(* IEC 61131-3 sources: Antarbhukti-LLM/DatasetCreation/SeedSTs/batch1_filtered_BASIC (part 2) *)

(* ---- FT_PROFILE.ST ---- *)
(*@PROPERTIES_EX@
TYPE: POU
LOCALE: 0
IEC_LANGUAGE: ST
PLC_TYPE: independent
PROC_TYPE: independent
GROUP: ENGINEERING.AUTOMATION
*)
(*@KEY@:DESCRIPTION*)
version 1.1	15 sep 2007
programmer 	tobias
tested by	hugo

FT_Profile generates an output signal which is defined by values over a time scale.
the different values are connected by ramps between the individual values.
a rising edge on E starts the output signal generation and E = True can delay time_3 / value_3 as long as it stays true.
an additional multiplier K can be used to multiply the output and an offset O can be added to the output dynamically.
(*@KEY@:END_DESCRIPTION*)
FUNCTION_BLOCK FT_PROFILE

(*Group:Default*)

VAR_INPUT
	K :	REAL := 1.0;
	O :	REAL := 0.0;
	M :	REAL := 1.0;
	E :	BOOL;
	VALUE_0 :	REAL;
	TIME_1 :	TIME;
	VALUE_1 :	REAL;
	TIME_2 :	TIME;
	VALUE_2 :	REAL;
	TIME_3 :	TIME;
	VALUE_3 :	REAL;
	TIME_10 :	TIME;
	VALUE_10 :	REAL;
	TIME_11 :	TIME;
	VALUE_11 :	REAL;
	TIME_12 :	TIME;
	VALUE_12 :	REAL;
	TIME_13 :	TIME;
	VALUE_13 :	REAL;
END_VAR

VAR_OUTPUT
	Y :	REAL;
	RUN :	BOOL;
	ET :	TIME;
END_VAR

VAR
	tx :	TIME;
	edge :	BOOL;
	state :	INT;
	ta :	TIME;
	tb :	TIME;
	t0 :	TIME;
	temp :	REAL;
	va :	REAL;
	vb :	REAL;
	T_PLC_MS :	T_PLC_MS;
END_VAR

(*@KEY@: WORKSHEET
NAME: FT_PROFILE
IEC_LANGUAGE: ST
*)
(* read system time *)
T_PLC_MS();
tx:= UDINT_TO_TIME(T_PLC_MS.T_PLC_MS);

(* determine start condition *)
IF E AND NOT edge THEN
	RUN := TRUE;
	ET := t#0s;
	t0 := tx;
	ta := tx;
	tb := multime(time_1, M);
	va := value_0;
	vb := value_1;
	temp := value_0;
	state := 1;
END_IF;
edge := E;

(* generate startup profile *)
IF run THEN
	CASE state OF
		1:	IF tx - ta >= tb THEN
				ta := ta + tb;
				tb := multime(time_2 - time_1, M);
				va := value_1;
				vb := value_2;
				temp := value_1;
				state := 2;
			ELSE
				temp := ((vb - va) * TIME_TO_REAL(tx - ta) / TIME_TO_REAL(tb) + va);
			END_IF;
		2:	IF tx - ta >= tb THEN
				ta := ta + tb;
				tb := multime(time_3 - time_2, M);
				va := value_2;
				vb := value_3;
				temp := value_2;
				state := 3;
			ELSE
				temp := ((vb - va) * TIME_TO_REAL(tx - ta) / TIME_TO_REAL(tb) + va);
			END_IF;
		3:	IF tx - ta >= tb THEN
				ta := ta + tb;
				tb := multime(time_10 - time_3, M);
				va := value_3;
				vb := value_10;
				temp := value_3;
				state := 4;
			ELSE
				temp := ((vb - va) * TIME_TO_REAL(tx - ta) / TIME_TO_REAL(tb) + va);
			END_IF;
		4 :	IF tx - ta >= tb THEN
				ta := ta + tb;
				tb := multime(time_11 - time_10, M);
				va := value_10;
				vb := value_11;
				temp := value_10;
				IF E THEN state := 5; ELSE state := 6; END_IF;
			ELSE
				temp := ((vb - va) * TIME_TO_REAL(tx - ta) / TIME_TO_REAL(tb) + va);
			END_IF;
		5:	(* extend the signal while E is true *)
			IF E THEN
				ta := tx;
			ELSE
				state := 6;
			END_IF;
		6:	IF tx - ta >= tb THEN
				ta := ta + tb;
				tb := multime(time_12 - time_11, M);
				va := value_11;
				vb := value_12;
				temp := value_11;
				state := 7;
			ELSE
				temp := ((vb - va) * TIME_TO_REAL(tx - ta) / TIME_TO_REAL(tb) + va);
			END_IF;
		7:	IF tx - ta >= tb THEN
				ta := ta + tb;
				tb := multime(time_13 - time_12, M);
				va := value_12;
				vb := value_13;
				temp := value_12;
				state := 8;
			ELSE
				temp := ((vb - va) * TIME_TO_REAL(tx - ta) / TIME_TO_REAL(tb) + va);
			END_IF;
		8:	IF tx - ta >= tb THEN
				temp := value_13;
				run := FALSE;
			ELSE
				temp := ((vb - va) * TIME_TO_REAL(tx - ta) / TIME_TO_REAL(tb) + va);
			END_IF;
	END_CASE;
	Y := temp * K + O;
	ET := tx - t0;
END_IF;

(* revision history
hm	27 feb 2007		rev 1.0
	original version

hm	15. sep2007		rev 1.1
	replaced Time() with T_PLC_MS for compatibility and performance reasons

*)
(*@KEY@: END_WORKSHEET *)
END_FUNCTION_BLOCK

(* ---- FT_PT1.ST ---- *)
(*@PROPERTIES_EX@
TYPE: POU
LOCALE: 0
IEC_LANGUAGE: ST
PLC_TYPE: independent
PROC_TYPE: independent
GROUP: ENGINEERING.CONTROL
*)
(*@KEY@:DESCRIPTION*)
version 1.11	18. jan. 2011
programmer 		hugo
tested by		oscat

FT_PT1 is an low pass filter with a programmable time T and faktor K.

(*@KEY@:END_DESCRIPTION*)
FUNCTION_BLOCK FT_PT1

(*Group:Default*)

VAR_INPUT
	IN :	REAL;
	T :	TIME;
	K :	REAL := 1.0;
END_VAR

VAR_OUTPUT
	OUT :	REAL;
END_VAR

VAR
	last :	UDINT;
	tx :	UDINT;
	init :	BOOL;
	T_PLC_US :	T_PLC_US;
END_VAR

(*@KEY@: WORKSHEET
NAME: FT_PT1
IEC_LANGUAGE: ST
*)
(* read system time *)
T_PLC_US();
tx:= T_PLC_US.T_PLC_US;

(* startup initialisation *)
IF NOT init OR T = t#0s THEN
	init := TRUE;
	out := K * in;
ELSE
	out := out + (in * K - out) * UDINT_TO_REAL(Tx - last) / TIME_TO_REAL(T) * 1.0E-3;
	IF ABS(out) < 1.0E-20 THEN out := 0.0; END_IF;
END_IF;
last := tx;

(*
hm 1.1.2007	rev 1.1
	corrected error while startup value was not correct
	for very small time values real output would run out of range.

hm 3.1.2007	rev 1.2
	corrected an error for falling edge failures.
	added output faktor K.

hm 27. 2. 2007	rev 1.3
	output will be input during init for definitive startup condition.

hm	15.9.2007	rev 1.4
	changed time() to T_PLC_US() for compatibilitxy resons
	increased internal accuracy to Microseconds instead of Milliseconds

hm	23. oct 2007	rev 1.5
	added out := in to the init statements

hm	30. nov 2007	rev 1.6
	changed out to be K * in during initialization

hm	5. jan 2008	rev 1.7
	improved code for better performance

hm	16. mar. 2008	rev 1.8
	added type conversion to avoid warning under codesys 3.0

hm	14. jun. 2008	rev 1.9
	improved code

hm	11. mar. 2009	rev 1.10
	real constants updated to new systax using dot

hm	18. jan. 2011	rev 1.11
	avoid underrun of out
*)
(*@KEY@: END_WORKSHEET *)
END_FUNCTION_BLOCK

(* ---- FT_PT2.ST ---- *)
(*@PROPERTIES_EX@
TYPE: POU
LOCALE: 0
IEC_LANGUAGE: ST
PLC_TYPE: independent
PROC_TYPE: independent
GROUP: ENGINEERING.CONTROL
*)
(*@KEY@:DESCRIPTION*)
version 1.5	11. mar. 2009
programmer 	hugo
tested by	oscat

FT_PT2 is a 2nd grade filter with programmable times T, D and faktor K.
(*@KEY@:END_DESCRIPTION*)
FUNCTION_BLOCK FT_PT2

(*Group:Default*)

VAR_INPUT
	IN :	REAL;
	T :	TIME;
	D :	REAL;
	K :	REAL := 1.0;
END_VAR

VAR_OUTPUT
	OUT :	REAL;
END_VAR

VAR
	init :	BOOL;
	int1 :	INTEGRATE;
	int2 :	INTEGRATE;
	tn :	REAL;
	I1 :	REAL;
	I2 :	REAL;
	tn2 :	REAL;
END_VAR

(*@KEY@: WORKSHEET
NAME: FT_PT2
IEC_LANGUAGE: ST
*)
(* startup initialisation *)
IF NOT init OR T = T#0s THEN
	init := TRUE;
	out := K * in;
	I2 := out;
ELSE
	TN := TIME_TO_REAL(T) / 1000.0;
	tn2 := TN * TN;
	int1(X := in * K / tn2 - I1 * 0.5 * D / TN - I2 / TN2, Y := I1);
	I1 := int1.Y;
	int2(X := I1,Y := I2);
	I2 := int2.Y;
	out := I2;
END_IF;

(* revision history

15.1.2007 hm		rev 1.1
	changed formula to new more acurate formula

hm 15.9.2007		rev 1.2
	deleted unused code for init system time reading tx

hm	30.11.2007	rev 1.3
	changed out to be K * in during initialization
	avoind divide by 0 if tn = 0

hm	3. nov. 2008	rev 1.4
	optimized code and fixed a problem with init

hm	11. mar. 2009	rev 1.5
	real constants updated to new systax using dot

*)
(*@KEY@: END_WORKSHEET *)
END_FUNCTION_BLOCK

(* ---- FT_RMP.ST ---- *)
(*@PROPERTIES_EX@
TYPE: POU
LOCALE: 0
IEC_LANGUAGE: ST
PLC_TYPE: independent
PROC_TYPE: independent
GROUP: MATHEMATICAL.FUNCTIONS
*)
(*@KEY@:DESCRIPTION*)
version 1.4	25 jan 2008
programmer 	oscat
tested BY	oscat

this ramp function follows an input signal with a linear ramp up or down, the up or down speed can be set with KF and KR.
a K factor of 1 means 1 unit per second on the output. K factors can only be positive and not negative.
a busy output signals the ramp is running or busy false means the in value is present on the output.
a rmp input false means the output follows the input dierctly while a rmp = true means the output follows the input with a ramp.
a updn output signal the directon of the ramp (up or down).
(*@KEY@:END_DESCRIPTION*)
FUNCTION_BLOCK FT_RMP

(*Group:Default*)

VAR_INPUT
	RMP :	BOOL := TRUE;
	IN :	REAL;
	KR :	REAL;
	KF :	REAL;
END_VAR

VAR_OUTPUT
	OUT :	REAL;
	BUSY :	BOOL;
	UD :	BOOL;
END_VAR

VAR
	tx :	TIME;
	last :	TIME;
	init :	BOOL;
	T_PLC_MS :	T_PLC_MS;
END_VAR

(*@KEY@: WORKSHEET
NAME: FT_RMP
IEC_LANGUAGE: ST
*)
(* read system time *)
T_PLC_MS();
tx:= UDINT_TO_TIME(T_PLC_MS.T_PLC_MS) - last;

IF NOT init THEN
	init := TRUE;
	last := tx;
	tx := t#0s;
	out := in;
END_IF;
IF NOT rmp THEN
	out := in;
	busy := FALSE;
ELSIF out > in THEN
	(* ramp down *)
	out := out - TIME_TO_REAL(tx) * 0.001 * KF;
	out := MAX(in, out);
ELSIF out < in THEN
	(* ramp up *)
	out := out + TIME_TO_REAL(tx) * 0.001 * KR;
	out := MIN(in, out);
END_IF;

(* set busy and dir flags *)
IF out < in THEN
	busy := TRUE;
	ud := TRUE;
ELSIF out > in THEN
	busy := TRUE;
	ud := FALSE;
ELSE
	busy := FALSE;
END_IF;
last := last + tx;

(* revision history:

hm 8.10.2006			rev 1.1
	added ud output

hm 12. feb 2007		rev 1.2
	added init variable and corrected a possible startup problem

hm	17. sep 2007	rev 1.3
	replaced time() with t_plc_ms() for compatibility reasons

hm	25. jan 2008	rev 1.4
	performance improvements
	allow KR and KF to be 0
*)
(*@KEY@: END_WORKSHEET *)
END_FUNCTION_BLOCK

(* ---- GEN_PULSE.ST ---- *)
(*@PROPERTIES_EX@
TYPE: POU
LOCALE: 0
IEC_LANGUAGE: ST
PLC_TYPE: independent
PROC_TYPE: independent
GROUP: ENGINEERING.SIGNAL_GENERATORS
*)
(*@KEY@:DESCRIPTION*)
version 1.5	8. apr. 2011
programmer 	hugo
tested by	oscat

GEN_PULSE uses the internal sps timer to generate a continuous output waveform with programmable high and low time.
the accuracy of gen_pulse is depending on the system timer.
when time is 0 the high and low times are exactly one cycle.
ENQ = TRUE will start and ENQ = FALSE will stop the generator.
(*@KEY@:END_DESCRIPTION*)
FUNCTION_BLOCK GEN_PULSE

(*Group:Default*)

VAR_INPUT
	ENQ :	BOOL := TRUE;
	PTH :	TIME;
	PTL :	TIME;
END_VAR

VAR_OUTPUT
	Q :	BOOL;
END_VAR

VAR
	T_PLC_MS :	T_PLC_MS;
	tx :	TIME;
	tn :	TIME;
	init :	BOOL;
END_VAR

(*@KEY@: WORKSHEET
NAME: GEN_PULSE
IEC_LANGUAGE: ST
*)
IF enq THEN
	T_PLC_MS();	(* read system timer *)
	tx:= UDINT_TO_TIME(T_PLC_MS.T_PLC_MS);
	IF NOT init THEN init := TRUE; tn := tx; END_IF;
	IF tx - tn >= SEL(Q, PTL, PTH) THEN
		tn := tn + SEL(Q, PTL, PTH);
		Q := NOT Q;
	END_IF;
ELSE
	Q := FALSE;
	init := FALSE;
END_IF;

(* revision history
hm	29. jun. 2008	rev 1.0
	original version

hm	23. nov. 2008	rev 1.1
	set default for enq to be true

hm	18. jul. 2009	rev 1.2
	improved performance

hm	13. nov. 2009	rev 1.3
	corrected error

hm	16. feb. 2011	rev 1.4
	corrected an error when timer overflows

hm	8. apr. 2011	rev 1.5
	ptl and pth was exchanged
*)
(*@KEY@: END_WORKSHEET *)
END_FUNCTION_BLOCK

(* ---- GEN_RMP.ST ---- *)
(*@PROPERTIES_EX@
TYPE: POU
LOCALE: 0
IEC_LANGUAGE: ST
PLC_TYPE: independent
PROC_TYPE: independent
GROUP: ENGINEERING.SIGNAL_GENERATORS
*)
(*@KEY@:DESCRIPTION*)
version 1.4	10. mar. 2009
programmer 	oscat
tested BY	oscat

this signal generator generates a ramp wave output. The ramp wave signal is defined by period time (PT),
amplitude (AM), offset (OS) and a specific delay for the output signal (DL).
The Output waveform will have its minimum peak at OS and its maximum peak at AM + OS.
The delay input can delay a signal up to PT, this can be useful to synchronize different generators
and generate interleaving signals.
in addition to the analog output Out there is a second boolean output Q with is true for one cycle when the ramp starts.

(*@KEY@:END_DESCRIPTION*)
FUNCTION_BLOCK GEN_RMP

(*Group:Default*)

VAR_INPUT
	PT :	TIME := T#1s;
	AM :	REAL := REAL#1.0;
	OS :	REAL;
	DL :	REAL;
END_VAR

VAR_OUTPUT
	Q :	BOOL;
	OUT :	REAL;
END_VAR

VAR
	tx :	TIME;
	last :	TIME;
	init :	BOOL;
	temp :	REAL;
	ltemp :	REAL;
	T_PLC_MS :	T_PLC_MS;
END_VAR

(*@KEY@: WORKSHEET
NAME: GEN_RMP
IEC_LANGUAGE: ST
*)
(* read system time and prepare input data *)
T_PLC_MS();
tx:= UDINT_TO_TIME(T_PLC_MS.T_PLC_MS) - last;
DL := modR(dl,1.0);
IF dl < 0.0 THEN dl := 1.0 - dl; END_IF;

(* init section *)
IF NOT init THEN
	init := TRUE;
	last := tx;
	tx := t#0s;
END_IF;

(* add last if one cycle is finished *)
IF tx >= pt THEN
	last := last + pt;
	tx := tx - pt;
END_IF;

(* generate sine wave *)
ltemp := temp;
IF pt > t#0s THEN temp := fract(TIME_TO_REAL(tx + multime(pt, dl)) / TIME_TO_REAL(pt)); END_IF;
out := am * temp + os;

(* boolean output Q *)
Q := temp < ltemp;

(* revision history
hm	3. mar 2007		rev 1.0
	original version

hm	17 sep 2007		rev 1.1
	replaced time() with t_plc_ms for compatibilitx reasons

hm	27. nov 2007	rev 1.2
	avoid divide by 0 when pt = 0

ks	26. oct. 2008	rev 1.3
	code optimization

hm	10. mar. 2009	rev 1.4
	changed real constants to use dot syntax
*)
(*@KEY@: END_WORKSHEET *)
END_FUNCTION_BLOCK

(* ---- GEN_SQ.ST ---- *)
(*@PROPERTIES_EX@
TYPE: POU
LOCALE: 0
IEC_LANGUAGE: ST
PLC_TYPE: independent
PROC_TYPE: independent
GROUP: LOGIC.GENERATORS
*)
(*@KEY@:DESCRIPTION*)
version 1.3	16. feb. 2011
programmer 	    hugo
tested by		tobias

gen_sq generates square wave signal with programmable period time.

(*@KEY@:END_DESCRIPTION*)
FUNCTION_BLOCK GEN_SQ

(*Group:Default*)

VAR_INPUT
	PT :	TIME;
END_VAR

VAR_OUTPUT
	Q :	BOOL;
END_VAR

VAR
	init :	BOOL;
	tn :	TIME;
	tx :	TIME;
	T_PLC_MS :	T_PLC_MS;
END_VAR

(*@KEY@: WORKSHEET
NAME: GEN_SQ
IEC_LANGUAGE: ST
*)
(* read system time *)
T_PLC_MS();
tx := UDINT_TO_TIME(T_PLC_MS.T_PLC_MS);

IF NOT init THEN
	init := TRUE;
	tn := tx;
	Q := TRUE;
ELSIF tx - tn >= DWORD_TO_TIME(SHR(TIME_TO_DWORD(PT),1)) THEN
	Q := NOT Q;
	tn := tn + DWORD_TO_TIME(SHR(TIME_TO_DWORD(pt),1));
END_IF;

(* revision history
hm	4. aug 2006	rev 1.0
	original version

hm	17. sep 2007	rev 1.1
	replaced time() with T_PLC_MS() for compatibility reasons

hm	18. jul. 2009	rev 1.2
	improved accuracy

hm	16. feb 2011	rev 1.3
	corrected an error with timer overflow
*)

(*@KEY@: END_WORKSHEET *)
END_FUNCTION_BLOCK

(* ---- HYST.ST ---- *)
(*@PROPERTIES_EX@
TYPE: POU
LOCALE: 0
IEC_LANGUAGE: ST
PLC_TYPE: independent
PROC_TYPE: independent
GROUP: ENGINEERING.CONTROL
*)
(*@KEY@:DESCRIPTION*)
version 1.0	2. jun. 2008
programmer 	hugo
tested BY	tobias

This Hystereses function has two modes:
1. if on > off then Q will be switched high when in > on and switched low when in < off.
2. if on < off then Q will be switched high when in < on and switched low when in > off.
the output win will be high when in is between low and high.
(*@KEY@:END_DESCRIPTION*)
FUNCTION_BLOCK HYST

(*Group:Default*)

VAR_INPUT
	IN :	REAL;
	ON :	REAL;
	OFF :	REAL;
END_VAR

VAR_OUTPUT
	Q :	BOOL;
	WIN :	BOOL;
END_VAR

(*@KEY@: WORKSHEET
NAME: HYST
IEC_LANGUAGE: ST
*)
IF ON >= OFF THEN
	IF IN < OFF THEN
		Q := FALSE;
		WIN := FALSE;
	ELSIF  IN > ON THEN
		Q := TRUE;
		WIN := FALSE;
	ELSE
		WIN := TRUE;
	END_IF;
ELSE
	IF IN > OFF THEN
		Q := FALSE;
		WIN := FALSE;
	ELSIF  IN < ON THEN
		Q := TRUE;
		WIN := FALSE;
	ELSE
		WIN := TRUE;
	END_IF;
END_IF;

(* revision history
hm		2.  jun 2008	rev 1.0
	original version

*)
(*@KEY@: END_WORKSHEET *)
END_FUNCTION_BLOCK

(* ---- HYST_1.ST ---- *)
(*@PROPERTIES_EX@
TYPE: POU
LOCALE: 0
IEC_LANGUAGE: ST
PLC_TYPE: independent
PROC_TYPE: independent
GROUP: ENGINEERING.CONTROL
*)
(*@KEY@:DESCRIPTION*)
version 1.1	2. jun. 2008
programmer 	hugo
tested BY	tobias

this hysteresis function switches the output high if the input signal reaches obove high and will switch to low when the input falls back below low value.
a separate output mid is set if the input stays between low and high value.
(*@KEY@:END_DESCRIPTION*)
FUNCTION_BLOCK HYST_1

(*Group:Default*)

VAR_INPUT
	IN :	REAL;
	HIGH :	REAL;
	LOW :	REAL;
END_VAR

VAR_OUTPUT
	Q :	BOOL;
	WIN :	BOOL;
END_VAR

(*@KEY@: WORKSHEET
NAME: HYST_1
IEC_LANGUAGE: ST
*)
IF in < low THEN
	Q := FALSE;
	win := FALSE;
ELSIF in > high THEN
	Q := TRUE;
	win := FALSE;
ELSE
	win := TRUE;
END_IF;

(* code used for rev 1.0
IF Q THEN
	IF in < low THEN q := FALSE; END_IF;
ELSE
	IF in > high THEN q := TRUE; END_IF;
END_IF;
win := in > low AND in < high;
*)
(*@KEY@: END_WORKSHEET *)
END_FUNCTION_BLOCK

(* ---- HYST_2.ST ---- *)
(*@PROPERTIES_EX@
TYPE: POU
LOCALE: 0
IEC_LANGUAGE: ST
PLC_TYPE: independent
PROC_TYPE: independent
GROUP: ENGINEERING.CONTROL
*)
(*@KEY@:DESCRIPTION*)
version 1.2	2. jun. 2008
programmer 	oscat
tested BY	tobias

this hysteresis function switches the output high if the input signal reaches obove val + hys/2 and will switch to low when the input falls back below val - hys/2 value.
a separate output mid is set if the input stays between low and high value.
(*@KEY@:END_DESCRIPTION*)
FUNCTION_BLOCK HYST_2

(*Group:Default*)

VAR_INPUT
	IN :	REAL;
	VAL :	REAL;
	HYS :	REAL;
END_VAR

VAR_OUTPUT
	Q :	BOOL;
	WIN :	BOOL;
END_VAR

VAR
	tmp :	REAL;
END_VAR

(*@KEY@: WORKSHEET
NAME: HYST_2
IEC_LANGUAGE: ST
*)
tmp := val - hys * 0.5;
IF in < tmp THEN
	Q := FALSE;
	win := FALSE;
ELSIF in > tmp + hys THEN
	Q := TRUE;
	win := FALSE;
ELSE
	win := TRUE;
END_IF;

(* code used for 1.2 and before
X := hys * 0.5;
IF Q THEN
	IF in < val - x THEN q := FALSE; END_IF;
ELSE
	IF in > val + x THEN q := TRUE; END_IF;
END_IF;
win := in > val - x AND in < val + x;
*)

(* revision history
hm		4. aug 2006	rev 1.0
	original version

hm		5. jan 2008	rev 1.1
	improved code for better performance

hm		2. jun. 2008	rev 1.2
	improved performance
*)
(*@KEY@: END_WORKSHEET *)
END_FUNCTION_BLOCK

(* ---- HYST_3.ST ---- *)
(*@PROPERTIES_EX@
TYPE: POU
LOCALE: 0
IEC_LANGUAGE: ST
PLC_TYPE: independent
PROC_TYPE: independent
GROUP: ENGINEERING.CONTROL
*)
(*@KEY@:DESCRIPTION*)
version 1.2	5 jan 2008
programmer 	oscat
tested BY	tobias

this is a double hysteresis function. Out1 follows a hysteresis function defined by val1and hyst, while out 2 follows val2 and hyst.
if the input signal is between the two hysteresis switches (val1 and val2) then non of the outputs is active.
(*@KEY@:END_DESCRIPTION*)
FUNCTION_BLOCK HYST_3

(*Group:Default*)

VAR_INPUT
	IN :	REAL;
	HYST :	REAL;
	VAL1 :	REAL;
	VAL2 :	REAL;
END_VAR

VAR_OUTPUT
	Q1 :	BOOL;
	Q2 :	BOOL;
END_VAR

VAR
	X :	REAL;
END_VAR

(*@KEY@: WORKSHEET
NAME: HYST_3
IEC_LANGUAGE: ST
*)
X := hyst * 0.5;
IF in < val1 - X THEN
	q1 := TRUE;
ELSIF in > val1 + X THEN
	q1 := FALSE;
END_IF;
IF in < val2 - X THEN
	q2 := FALSE;
ELSIF in > val2 + X THEN
	q2 := TRUE;
END_IF;

(* revision history
hm	22. jan 2007	rev 1.0
	original version

hm	27. dec 2007	rev 1.1
	changed code for better performance

hm	5. jan 2008		rev 1.2
	further performance iprovements

*)
(*@KEY@: END_WORKSHEET *)
END_FUNCTION_BLOCK

(* ---- INC_DEC.ST ---- *)
(*@PROPERTIES_EX@
TYPE: POU
LOCALE: 0
IEC_LANGUAGE: ST
PLC_TYPE: independent
PROC_TYPE: independent
GROUP: ENGINEERING.AUTOMATION
*)
(*@KEY@:DESCRIPTION*)
version 1.0	4 aug 2006
programmer 	oscat
tested BY	oscat

incremental decoder with quadruple accuracy.
2 pulses for each channel are created for each directional pulse.
(*@KEY@:END_DESCRIPTION*)
FUNCTION_BLOCK INC_DEC

(*Group:Default*)

VAR_INPUT
	CHA :	BOOL;
	CHB :	BOOL;
	RST :	BOOL := 0;
END_VAR

VAR_OUTPUT
	DIR :	BOOL;
	CNT :	INT;
END_VAR

VAR
	edgea :	BOOL := 0;
	clk :	BOOL;
	clka :	BOOL;
	clkb :	BOOL;
	edgeb :	BOOL;
	axb :	BOOL;
END_VAR

(*@KEY@: WORKSHEET
NAME: INC_DEC
IEC_LANGUAGE: ST
*)
axb := cha XOR chb;

(* create pulses for channel a *)
clka := cha XOR edgea;
edgea := cha;

clkb := chb XOR edgeb;
edgeb := chb;

(* create pulses for both channels *)
clk := clka OR clkb;

(* set the direction output *)
IF axb AND clka THEN dir := TRUE; END_IF;
IF axb AND clkb THEN dir := FALSE; END_IF;

(* increment or decrement the counter *)
IF clk AND dir THEN cnt := cnt + 1; END_IF;
IF clk AND NOT dir THEN cnt := cnt -1; END_IF;

(* reset the counter if rst active *)
IF rst THEN cnt := 0; END_IF;
(*@KEY@: END_WORKSHEET *)
END_FUNCTION_BLOCK

(* ---- INTERLOCK.ST ---- *)
(*@PROPERTIES_EX@
TYPE: POU
LOCALE: 0
IEC_LANGUAGE: ST
PLC_TYPE: independent
PROC_TYPE: independent
GROUP: ENGINEERING.AUTOMATION
*)
(*@KEY@:DESCRIPTION*)
version 1.0	28 sep 2007
programmer 	hugo
tested by	tobias

INTERLOCK has two inputs I1 and I2 which drive the corresponding outputs Q1 and Q2.
the inputs signals lock each other out and therfore I1 can only drive Q1 when I2 is Low and vice versa.
The input TL specifies a dead time between two outputs can become active.
an output can only become active when the other output was not active for the time TL.
(*@KEY@:END_DESCRIPTION*)
FUNCTION_BLOCK INTERLOCK

(*Group:Default*)

VAR_INPUT
	I1 :	BOOL;
	I2 :	BOOL;
	TL :	TIME;
END_VAR

VAR_OUTPUT
	Q1 :	BOOL;
	Q2 :	BOOL;
END_VAR

VAR
	T1 :	TOF;
	T2 :	TOF;
END_VAR

(*@KEY@: WORKSHEET
NAME: INTERLOCK
IEC_LANGUAGE: ST
*)
(* the input signal have a run delay to lockout the other input *)
T1(IN := I1, PT := TL);
T2(IN := I2, PT := TL);

Q1 := I1 AND NOT t2.Q;
Q2 := I2 AND NOT t1.Q;

(* revision history

hm	28 sep 2007		rev 1.0
	original version

*)
(*@KEY@: END_WORKSHEET *)
END_FUNCTION_BLOCK

(* ---- INTERLOCK_4.ST ---- *)
(*@PROPERTIES_EX@
TYPE: POU
LOCALE: 0
IEC_LANGUAGE: ST
PLC_TYPE: independent
PROC_TYPE: independent
GROUP: ENGINEERING.AUTOMATION
*)
(*@KEY@:DESCRIPTION*)
version 1.1	14. mar. 2009
programmer 	hugo
tested by	oscat

INTERLOCK_4 detects one of 4 switches and delivers the number of the switch pressed on the output out
a output tp is true for one cycle if the output has changed.
a setup variable MODE selects between 3 different modes:
MODE = 0, any input active will disable all other inputs
MODE = 1, the input with the highest number will be acepted
mode = 2, the input last pressed will disable all others

(*@KEY@:END_DESCRIPTION*)
FUNCTION_BLOCK INTERLOCK_4

(*Group:Default*)

VAR_INPUT
	I0 :	BOOL;
	I1 :	BOOL;
	I2 :	BOOL;
	I3 :	BOOL;
	E :	BOOL;
	MODE :	INT;
END_VAR

VAR_OUTPUT
	OUT :	BYTE;
	TP :	BOOL;
END_VAR

VAR
	in :	BYTE;
	last :	BYTE;
	old :	BYTE;
	lmode :	INT;
END_VAR

(*@KEY@: WORKSHEET
NAME: INTERLOCK_4
IEC_LANGUAGE: ST
*)
(* check if enable is active *)
IF E THEN
(* reset all vars when there is a mode change on thy fly *)
	IF mode <> lmode THEN
		out := BYTE#0;
		last := BYTE#0;
		old := BYTE#0;
		lmode := mode;
	END_IF;
	(* load inputs into in *)
	in:=BIT_LOAD_B(in,I0,0); (* in.0 *)
	in:=BIT_LOAD_B(in,I1,1); (* in.1 *)
	in:=BIT_LOAD_B(in,I2,2); (* in.2 *)
	in:=BIT_LOAD_B(in,I3,3); (* in.3 *)
	(* only execute when there is any change *)
	IF in <> last THEN
		(* only execute when inputs have chages state *)
		CASE mode OF
			0:	(* output directly display inputs as bits in byte out *)
				out := in;

			1:	(* the input with the highest number will be acepted *)
				IF    (in AND BYTE#2#00001000) > BYTE#0 (* in.3 *) THEN out := BYTE#8;
				ELSIF (in AND BYTE#2#00000100) > BYTE#0 (* in.2 *) THEN out := BYTE#4;
				ELSIF (in AND BYTE#2#00000010) > BYTE#0 (* in.1 *) THEN out := BYTE#2;
				ELSE out := in;
				END_IF;

			2:	(* input last pressed will be displayed only *)
				last := ((in XOR last) AND in);
				IF    (last AND BYTE#2#00001000) > BYTE#0 (* last.3 *) THEN out := BYTE#8;
				ELSIF (last AND BYTE#2#00000100) > BYTE#0 (* last.2 *) THEN out := BYTE#4;
				ELSIF (last AND BYTE#2#00000010) > BYTE#0 (* last.1 *) THEN out := BYTE#2;
				ELSE out := last;
				END_IF;

			3:	(* any input active will disable all other inputs *)
				IF (out AND in) = BYTE#0 THEN
					IF    (in AND BYTE#2#00001000) > BYTE#0 (* in.3 *) THEN out := BYTE#8;
					ELSIF (in AND BYTE#2#00000100) > BYTE#0 (* in.2 *) THEN out := BYTE#4;
					ELSIF (in AND BYTE#2#00000010) > BYTE#0 (* in.1 *) THEN out := BYTE#2;
					ELSE out := in;
					END_IF;
				END_IF;

		END_CASE;
		last := in;
	END_IF;
	tp := out <> old;
	old := out;
ELSE
	out := BYTE#0;
	last := BYTE#0;
	old := BYTE#0;
	lmode := 0;
	tp := FALSE;
END_IF;

(* revision history
hm	24. oct 2008	rev 1.0
	original version

hm	14. mar. 2009	rev 1.1
	replaced double assignments

*)
(*@KEY@: END_WORKSHEET *)
END_FUNCTION_BLOCK

(* ---- LTCH.ST ---- *)
(*@PROPERTIES_EX@
TYPE: POU
LOCALE: 0
IEC_LANGUAGE: ST
PLC_TYPE: independent
PROC_TYPE: independent
GROUP: LOGIC.FF_PULSE_TRIGGERED
*)
(*@KEY@:DESCRIPTION*)
version 1.2	30. oct. 2008
programmer 	hugo
tested by	oscat

Transparent Latch with asynchronous reset
(*@KEY@:END_DESCRIPTION*)
FUNCTION_BLOCK LTCH

(*Group:Default*)

VAR_INPUT
	D :	BOOL;
	L :	BOOL;
	RST :	BOOL;
END_VAR

VAR_OUTPUT
	Q :	BOOL;
END_VAR

(*@KEY@: WORKSHEET
NAME: LTCH
IEC_LANGUAGE: ST
*)
(* as long as L is true, the latch is transparent and and change of D is transferred to Q *)
(* of course only when there is no asynchronous reset *)
IF rst THEN				(* if asynchronous reset then Q=0 *)
	Q := FALSE;
ELSIF L THEN			(* latch is transparent *)
	Q := D;
END_IF;

(* revision history
hm	4. aug 2006		rev 1.0
	original version

hm	27. dec 2007	rev 1.1
	changed code for better performance

hm	30. oct. 2008	rev 1.2
	deleted unnecessary init with 0

*)
(*@KEY@: END_WORKSHEET *)
END_FUNCTION_BLOCK

(* ---- LTCH_4.ST ---- *)
(*@PROPERTIES_EX@
TYPE: POU
LOCALE: 0
IEC_LANGUAGE: ST
PLC_TYPE: independent
PROC_TYPE: independent
GROUP: LOGIC.FF_PULSE_TRIGGERED
*)
(*@KEY@:DESCRIPTION*)
version 1.3	14. mar. 2009
programmer 	hugo
tested by	oscat

Quad Transparent Latch with asynchronous reset
(*@KEY@:END_DESCRIPTION*)
FUNCTION_BLOCK LTCH_4

(*Group:Default*)

VAR_INPUT
	D0 :	BOOL;
	D1 :	BOOL;
	D2 :	BOOL;
	D3 :	BOOL;
	L :	BOOL;
	RST :	BOOL;
END_VAR

VAR_OUTPUT
	Q0 :	BOOL;
	Q1 :	BOOL;
	Q2 :	BOOL;
	Q3 :	BOOL;
END_VAR

(*@KEY@: WORKSHEET
NAME: LTCH_4
IEC_LANGUAGE: ST
*)
(* as long as L is true, the latch is transparent and and change of D is transferred to Q *)
(* of course only when there is no asynchronous reset *)
IF rst THEN			(* if asynchronous reset then Q=0 *)
	Q0 := FALSE;
	Q1 := FALSE;
	Q2 := FALSE;
	Q3 := FALSE;
ELSIF L THEN			(* latch is transparent *)
	Q0 := D0;
	Q1 := D1;
	Q2 := D2;
	Q3 := D3;
END_IF;

(* revision history
hm	4. aug 2006	rev 1.0
	original version

hm	27. dec 2007	rev 1.1
	changed code for better performance

hm	30. oct. 2008	rev 1.2
	deleted unnecessary init with 0

hm	14. mar. 2009	rev 1.3
	removed double assignments

*)
(*@KEY@: END_WORKSHEET *)
END_FUNCTION_BLOCK

(* ---- MANUAL_1.ST ---- *)
(*@PROPERTIES_EX@
TYPE: POU
LOCALE: 0
IEC_LANGUAGE: ST
PLC_TYPE: independent
PROC_TYPE: independent
GROUP: ENGINEERING.AUTOMATION
*)
(*@KEY@:DESCRIPTION*)
version 1.2	14. mar. 2009
programmer 	hugo
tested by	oscat

MANUAL_1 is a manual override for digital signals.
When MAN = FALSE, the output follows IN and when MAN = TRUE the Output follows M_I.

(*@KEY@:END_DESCRIPTION*)
FUNCTION_BLOCK MANUAL_1

(*Group:Default*)

VAR_INPUT
	IN :	BOOL;
	MAN :	BOOL;
	M_I :	BOOL;
	SET :	BOOL;
	RST :	BOOL;
END_VAR

VAR_OUTPUT
	Q :	BOOL;
	STATUS :	BYTE;
END_VAR

VAR
	S_edge :	BOOL;
	r_edge :	BOOL;
	edge :	BOOL;
END_VAR

(*@KEY@: WORKSHEET
NAME: MANUAL_1
IEC_LANGUAGE: ST
*)
IF NOT man THEN
	Q := IN;
	STATUS := BYTE#100;
	edge := FALSE;
ELSIF NOT s_edge AND set THEN
	Q := TRUE;
	edge := TRUE;
	status := BYTE#101;
ELSIF NOT r_edge AND rst THEN
	Q := FALSE;
	edge := TRUE;
	status := BYTE#102;
ELSIF NOT edge THEN
	Q := M_I;
	status := BYTE#103;
END_IF;

(* remember levels of manual signals *)
s_edge := SET;
r_edge := RST;

(* revision history
hm	17. jun 2008	rev 1.0
	original version

hm	17. oct 2008	rev 1.1
	deleted unnecessary variable m_edge

hm	14. mar. 2009	rev 1.2
	replaced double assignments

*)
(*@KEY@: END_WORKSHEET *)
END_FUNCTION_BLOCK

(* ---- MANUAL_2.ST ---- *)
(*@PROPERTIES_EX@
TYPE: POU
LOCALE: 0
IEC_LANGUAGE: ST
PLC_TYPE: independent
PROC_TYPE: independent
GROUP: ENGINEERING.AUTOMATION
*)
(*@KEY@:DESCRIPTION*)
version 1.0	22. sep. 2008
programmer 	hugo
tested by	oscat

MANUAL_2 is a manual override for boolean signals.
it has static force high and low as well as a manual input.
(*@KEY@:END_DESCRIPTION*)
FUNCTION_BLOCK MANUAL_2

(*Group:Default*)

VAR_INPUT
	IN :	BOOL;
	ENA :	BOOL;
	ON :	BOOL;
	OFF :	BOOL;
	MAN :	BOOL;
END_VAR

VAR_OUTPUT
	Q :	BOOL;
	STATUS :	BYTE;
END_VAR

(*@KEY@: WORKSHEET
NAME: MANUAL_2
IEC_LANGUAGE: ST
*)
IF ena THEN
	IF NOT ON AND NOT OFF THEN
		Q := IN;
		STATUS := BYTE#100;
	ELSIF on AND NOT off THEN
		Q := TRUE;
		STATUS := BYTE#101;
	ELSIF NOT on AND off THEN
		q := FALSE;
		STATUS := BYTE#102;
	ELSE
		Q := MAN;
		STATUS := BYTE#103;
	END_IF;
ELSE
	Q := FALSE;
	STATUS := BYTE#104;
END_IF;

(* revision history
hm	22. sep. 2008		rev 1.0
	original version

*)
(*@KEY@: END_WORKSHEET *)
END_FUNCTION_BLOCK

(* ---- MANUAL_4.ST ---- *)
(*@PROPERTIES_EX@
TYPE: POU
LOCALE: 0
IEC_LANGUAGE: ST
PLC_TYPE: independent
PROC_TYPE: independent
GROUP: ENGINEERING.AUTOMATION
*)
(*@KEY@:DESCRIPTION*)
version 1.0	17. jun 2008
programmer 	hugo
tested by	oscat

MANUAL_4 is a manual override for digital signals.
When MAN = FALSE, the output follows IN and when MAN = TRUE the Output follows M_I.
(*@KEY@:END_DESCRIPTION*)
FUNCTION_BLOCK MANUAL_4

(*Group:Default*)

VAR_INPUT
	I0 :	BOOL;
	I1 :	BOOL;
	I2 :	BOOL;
	I3 :	BOOL;
	MAN :	BOOL;
	STP :	BOOL;
	M0 :	BOOL;
	M1 :	BOOL;
	M2 :	BOOL;
	M3 :	BOOL;
END_VAR

VAR_OUTPUT
	Q0 :	BOOL;
	Q1 :	BOOL;
	Q2 :	BOOL;
	Q3 :	BOOL;
	STATUS :	BYTE;
END_VAR

VAR
	edge :	BOOL;
	pos :	INT;
	tog :	BOOL;
END_VAR

(*@KEY@: WORKSHEET
NAME: MANUAL_4
IEC_LANGUAGE: ST
*)
IF man THEN
	IF NOT TOG THEN
		Q0 := M0;
		Q1 := M1;
		Q2 := M2;
		Q3 := M3;
		STATUS := BYTE#101;
	END_IF;
	IF STP AND NOT edge THEN
		tog := TRUE;
		CASE pos OF
			0:	Q0 := TRUE;
				Q1 := FALSE;
				Q2 := FALSE;
				Q3 := FALSE;
				STATUS := BYTE#110;
			1:	Q0 := FALSE;
				Q1 := TRUE;
				Q2 := FALSE;
				Q3 := FALSE;
				STATUS := BYTE#111;
			2:	Q0 := FALSE;
				Q1 := FALSE;
				Q2 := TRUE;
				Q3 := FALSE;
				STATUS := BYTE#112;
			3:	Q0 := FALSE;
				Q1 := FALSE;
				Q2 := FALSE;
				Q3 := TRUE;
				STATUS := BYTE#113;
		END_CASE;
		pos := INC(pos,1,3);
	END_IF;
ELSE
	Q0 := I0;
	Q1 := I1;
	Q2 := I2;
	Q3 := I3;
	STATUS := BYTE#100;
	tog := FALSE;
	pos := 0;
END_IF;

(* remember status of stp *)
edge := STP;

(* revision history
hm	17. jun 2008		rev 1.0
	original version

*)
(*@KEY@: END_WORKSHEET *)
END_FUNCTION_BLOCK

(* ---- MESSAGE_4R.ST ---- *)
(*@PROPERTIES_EX@
TYPE: POU
LOCALE: 0
IEC_LANGUAGE: ST
PLC_TYPE: independent
PROC_TYPE: independent
GROUP: STRINGS
*)
(*@KEY@:DESCRIPTION*)
version 1.1	27. oct. 2008
programmer 	hugo
tested by	tobias

this function generates a rotation meassage with up to 4 strings.
on each rising edge of EN the next message in line will be displayed.
when EN stays high longer then one cycle, the next message will be displayed automatically after the time T1 is elapsed.
the output MX is the generated message and CX is a counter 0..3 signaling the current message displayed.
the displayed messages are 0 .. MM.
(*@KEY@:END_DESCRIPTION*)
FUNCTION_BLOCK MESSAGE_4R

(*Group:Default*)

VAR_INPUT
	M0 :	STRING;
	M1 :	STRING;
	M2 :	STRING;
	M3 :	STRING;
	MM :	INT := 3;
	ENQ :	BOOL := TRUE;
	CLK :	BOOL := TRUE;
	T1 :	TIME := T#3s;
END_VAR

VAR_OUTPUT
	MX :	STRING;
	MN :	INT;
	TR :	BOOL;
END_VAR

VAR
	timer :	TON;
	edge :	BOOL;
END_VAR

(*@KEY@: WORKSHEET
NAME: MESSAGE_4R
IEC_LANGUAGE: ST
*)
(* check for rising edge on EN *)
TR := FALSE;
IF ENQ THEN
	IF (NOT edge AND clk) OR timer.q THEN
			MN := INC1(MN, MM);
			TR := TRUE;
			timer(in := FALSE);
			CASE MN OF
				0 : MX := M0;
				1 : MX := M1;
				2 : MX := M2;
				3 : MX := M3;
			END_CASE;
	END_IF;
	edge := clk;
	timer( in := CLK, pt := T1);
ELSE
	MX := '';
	MN := 0;
END_IF;

(* revision history
hm	8. oct. 2008	rev 1.0
	original version

hm	27. oct. 2008	rev 1.1
	changed _INC to INC1

*)
(*@KEY@: END_WORKSHEET *)
END_FUNCTION_BLOCK

(* ---- MESSAGE_8.ST ---- *)
(*@PROPERTIES_EX@
TYPE: POU
LOCALE: 0
IEC_LANGUAGE: ST
PLC_TYPE: independent
PROC_TYPE: independent
GROUP: STRINGS
*)
(*@KEY@:DESCRIPTION*)
version 1.1	29. mar. 2008
programmer 	hugo
tested by	tobias

this function generates one out of 4 messages specified by S1 .. S8.
the selected message will be presented at the output M.
In1 has higher priority then In2 which has higher priority then IN3 and in8 has the lowest priority.
(*@KEY@:END_DESCRIPTION*)
FUNCTION_BLOCK MESSAGE_8

(*Group:Default*)

VAR_INPUT
	IN1 :	BOOL;
	IN2 :	BOOL;
	IN3 :	BOOL;
	IN4 :	BOOL;
	IN5 :	BOOL;
	IN6 :	BOOL;
	IN7 :	BOOL;
	IN8 :	BOOL;
	S1 :	STRING;
	S2 :	STRING;
	S3 :	STRING;
	S4 :	STRING;
	S5 :	STRING;
	S6 :	STRING;
	S7 :	STRING;
	S8 :	STRING;
END_VAR

VAR_OUTPUT
	M :	STRING;
END_VAR

(*@KEY@: WORKSHEET
NAME: MESSAGE_8
IEC_LANGUAGE: ST
*)
(* check if an alarm is present if yes set the output M otherwise clear M *)
IF in1 THEN
	M := S1;
ELSIF in2 THEN
	M := S2;
ELSIF in3 THEN
	M := S3;
ELSIF in4 THEN
	M := S4;
ELSIF in5 THEN
	M := S5;
ELSIF in6 THEN
	M := S6;
ELSIF in7 THEN
	M := S7;
ELSIF in8 THEN
	M := S8;
ELSE
	M := '';
END_IF;

(* revision history
hm	26.12.2007		rev 1.0
	original version

hm	29. mar. 2008	rev 1.1
	changed STRING to STRING(STRING_LENGTH)
*)
(*@KEY@: END_WORKSHEET *)
END_FUNCTION_BLOCK

(* ---- METER.ST ---- *)
(*@PROPERTIES_EX@
TYPE: POU
LOCALE: 0
IEC_LANGUAGE: ST
PLC_TYPE: independent
PROC_TYPE: independent
GROUP: ENGINEERING.MEASUREMENTS
*)
(*@KEY@:DESCRIPTION*)
version 1.4	8. mar. 2009
programmer 	oscat
tested BY	oscat

METER measures usage of power or similar values the output MX is the sum of the inputs over time.
MX := sum over time of (I1 * P1 + I2 * P2)/D.
a simple example is the consumption counter for a 2 stage oil burner where stage 1 is 10KW and stage 2 is 20KW.
I1 and I2 decide which value is accounted for, I1 = True only counts P1, I2 is True counts P2
and I1 and I2 is true counts P1 and P2.
the meter can be used for all kind of consumption meters. P1 and P2 can change on the fly.

(*@KEY@:END_DESCRIPTION*)
FUNCTION_BLOCK METER

(*Group:Default*)

VAR_INPUT
	M1 :	REAL;
	M2 :	REAL;
	I1 :	BOOL;
	I2 :	BOOL;
	D :	REAL := 1.0;
	RST :	BOOL;
END_VAR

VAR_IN_OUT
	MX :	REAL;
END_VAR

VAR RETAIN
	MR :	REAL2;
END_VAR

VAR
	MX1 :	REAL;(*current consumption value on M1 and M2*)
	MX2 :	REAL;(*current consumption value on M1 and M2*)
	tx :	UDINT;
	last :	UDINT;
	tc :	REAL;
	init :	BOOL;
	T_PLC_MS :	T_PLC_MS;
	R2_ADD :	R2_ADD;
END_VAR

(*@KEY@: WORKSHEET
NAME: METER
IEC_LANGUAGE: ST
*)
(* measure the last cycle time and make sure we onle execute once every millisecond *)
T_PLC_MS();
tx:= T_PLC_MS.T_PLC_MS;
IF NOT init THEN
	init := TRUE;
	last := tx;
	mr.RX := mx;
	mr.R1 := 0.0;
ELSIF tx = last THEN
	RETURN;
ELSE
	tc := UDINT_TO_REAL(tx - last) * 0.001;
END_IF;
last := tx;

(* reset *)
IF rst THEN
	mr.R1 := 0.0;
	mr.RX := 0.0;
ELSE
	(* current consumption measurement *)
	MX1 := SEL(I1,0.0,M1);
	MX2 := SEL(I2,0.0,M2);
	(* add up the current values in a double real *)
	R2_ADD(X:=MR,Y:=(SEL(I1,0.0,mx1) + SEL(I2, 0.0, mx2)) / D * TC);
	MR:=R2_ADD.R2_ADD;
	(* set the current output value *)
	MX := mr.RX;
END_IF;

(* revision history

hm	16. sep.2007		rev 1.0
	original version

hm	7. feb 2008		rev 1.1
	use new version of ft_int to avoid a counting stop at high values
	deleted unnecessary limits

hm	24. mar. 2008		rev 1.2
	use data_type real2 to extend accuracy to 15 digits total
	do not use ft_int which adds unnecessary overhead

hm	8. feb. 2009		rev 1.3
	changed mx to be I/O
	make sure calculation works for cycle times < 1 ms

hm	8. mar. 2009	rev 1.4
	last was not updated
	code improvements

*)

(*@KEY@: END_WORKSHEET *)
END_FUNCTION_BLOCK

(* ---- METER_STAT.ST ---- *)
(*@PROPERTIES_EX@
TYPE: POU
LOCALE: 0
IEC_LANGUAGE: ST
PLC_TYPE: independent
PROC_TYPE: independent
GROUP: ENGINEERING.MEASUREMENTS
*)
(*@KEY@:DESCRIPTION*)
version 1.3	18. jul. 2009
programmer 	oscat
tested BY	oscat

METER_STAT runs statistics of a metered value, it calculates the current week, day, month and year consumption and stores the corresponding last day, week, month and year value.

(*@KEY@:END_DESCRIPTION*)
FUNCTION_BLOCK METER_STAT

(*Group:Default*)

VAR_INPUT
	IN :	REAL;
	DI :	UDINT;
	RST :	BOOL;
END_VAR

VAR_IN_OUT
	LAST_DAY :	REAL;
	CURRENT_DAY :	REAL;
	LAST_WEEK :	REAL;
	CURRENT_WEEK :	REAL;
	LAST_MONTH :	REAL;
	CURRENT_MONTH :	REAL;
	LAST_YEAR :	REAL;
	CURRENT_YEAR :	REAL;
END_VAR

VAR RETAIN
	year_start :	REAL;
	month_start :	REAL;
	week_start :	REAL;
	day_start :	REAL;
	last_run :	UDINT;
END_VAR

(*@KEY@: WORKSHEET
NAME: METER_STAT
IEC_LANGUAGE: ST
*)
IF rst THEN
	Last_Day := 0.0;
	Current_Day := 0.0;
	Day_start := IN;
	Last_week := 0.0;
	Current_week := 0.0;
	Week_start := in;
	Last_month := 0.0;
	Current_month := 0.0;
	month_start := in;
	last_year := 0.0;
	current_year := 0.0;
	year_start := in;
ELSE
	Current_Day := IN - Day_Start;
	Current_Week := In - Week_Start;
	Current_Month := IN - Month_Start;
	Current_Year := IN - Year_Start;
END_IF;

IF YEAR_OF_DATE(DI) > YEAR_OF_DATE(last_run) THEN
	(* a new year has started *)
	last_year := current_year;
	current_year := 0.0;
	year_start := in;
	last_month := current_month;
	current_month := 0.0;
	month_start := in;
	last_day := current_day;
	current_day := 0.0;
	day_start := in;
ELSIF MONTH_OF_DATE(DI) > MONTH_OF_DATE(last_run) THEN
	(* a new month has started, january is alrerady done by year change *)
	last_month := current_month;
	current_month := 0.0;
	month_start := in;
	last_day := current_day;
	current_day := 0.0;
	day_start := in;
ELSIF DAY_OF_YEAR(di) > DAY_OF_YEAR(last_run) THEN
	(* day has chaged, first day of year and first day of month has already been taken care of *)
	last_day := current_day;
	current_day := 0.0;
	day_start := in;
END_IF;
IF DAY_OF_WEEK(DI) < DAY_OF_WEEK(last_run) THEN
	(* a new week has started *)
	last_week := current_week;
	current_week := 0.0;
	week_start := in;
END_IF;
last_run := di;

(* revision history
hm	16. sep. 2007	rev 1.0
	original version

hm	7. oct. 2008	rev 1.1
	changed function year_to_year_of_date
	changed function month to month_of_date
	changed function weekday to day_of_week

hm	11. mar. 2009	rev 1.2
	changed real constants to use dot syntax

hm	18. jul. 2009	rev 1.3
	changes all outputs to be I/O
*)

(*@KEY@: END_WORKSHEET *)
END_FUNCTION_BLOCK

(* ---- ONTIME.ST ---- *)
(*@PROPERTIES_EX@
TYPE: POU
LOCALE: 0
IEC_LANGUAGE: ST
PLC_TYPE: independent
PROC_TYPE: independent
GROUP: ENGINEERING.MEASUREMENTS
*)
(*@KEY@:DESCRIPTION*)
version 2.5	18. mar. 2011
programmer 	oscat
tested by	tobias

ONTIME measures the ontime of a signal in seconds.
the output SECONDS is of type DWORD which results in a total measurement range of 1 second up to 136 years.
internally ontime works with a resolution of milliseconds
(*@KEY@:END_DESCRIPTION*)
FUNCTION_BLOCK ONTIME

(*Group:Default*)

VAR_INPUT
	IN :	BOOL;
	RST :	BOOL;
END_VAR

VAR_IN_OUT
	SECONDS :	UDINT;
	CYCLES :	UDINT;
END_VAR

VAR
	tx :	UDINT;
	last :	UDINT;
	edge :	BOOL;
	init :	BOOL;
	ms :	UDINT;
	T_PLC_MS :	T_PLC_MS;
END_VAR

(*@KEY@: WORKSHEET
NAME: ONTIME
IEC_LANGUAGE: ST
*)
(* read system time *)
T_PLC_MS();
tx:= T_PLC_MS.T_PLC_MS;

(* make sure the first cycle works correctly *)
IF NOT init THEN
	init := TRUE;
	last := tx;
	ms := UDINT#0;
END_IF;
IF RST THEN
	SECONDS := UDINT#0;
	CYCLES := UDINT#0;
	last := tx;
	ms := UDINT#0;
ELSIF IN THEN
	(* add the current milliseconds *)
	ms := (tx - last) + ms;
	IF ms >= UDINT#1000 THEN
		seconds := seconds + UDINT#1;
		ms := ms - UDINT#1000;
	END_IF;
	cycles := cycles + BOOL_TO_UDINT(NOT edge);
END_IF;
last := tx;
edge := in;

(* revision history
hm 22.2.2007		rev 1.1
	changed VAR RETAIN PERSISTENT to VAR RETAIN for better compatibility
	wago lon contollers do not support persisitent

hm 2.8.2007		rev 1.2
	adding time up in a real number will automatically lead to the point where
	small time scales like the cycle time will be below the resolution of real and therefore
	ontime would not increase in small steps as necessary
	the time is now measured internally in two  dwords and be converted to real only for
	output purposes.
	deleted the variable power because it was unnecessary

hm	16.9.2007		rev 1.3
	changes time() to T_plc_ms() for compatibility reasons

hm	2. dec. 2007	rev 1.4
	chaged code for better performance

hm	16. mar. 2008	rev 1.5
	added type conversions to avoid warnings under codesys 3.0

hm	21. oct. 2008	rev 2.0
	changed module for much better performance and allow for external result storage

hm	10. nov. 2008	rev 2.1
	increased internal resolution to milliseconds

hm	16. nov. 2008	rev 2.2
	changed typecast to avoid warnings

hm	17. dec. 2008	rev 2.3
	fixed an error when in would be true for more then 49 days

hm	17. jan 2011	rev 2.4
	init will not clear seconds and cycles, only rst clears these values

hm	18. mar. 2011	rev 2.5
	reset was not working

*)

(*@KEY@: END_WORKSHEET *)
END_FUNCTION_BLOCK

(* ---- PWM_DC.ST ---- *)
(*@PROPERTIES_EX@
TYPE: POU
LOCALE: 0
IEC_LANGUAGE: ST
PLC_TYPE: independent
PROC_TYPE: independent
GROUP: ENGINEERING.SIGNAL_GENERATORS
*)
(*@KEY@:DESCRIPTION*)
version 1.4	11. mar. 2009
programmer 	oscat
tested BY	oscat

this signal generator generates a square wave signal which is specified by the frequency and the duty cycle

(*@KEY@:END_DESCRIPTION*)
FUNCTION_BLOCK PWM_DC

(*Group:Default*)

VAR_INPUT
	F :	REAL;
	DC :	REAL;
END_VAR

VAR_OUTPUT
	Q :	BOOL;
END_VAR

VAR
	clk :	CLK_Prg;
	pulse :	TP_X;
	tmp :	REAL;
END_VAR

(*@KEY@: WORKSHEET
NAME: PWM_DC
IEC_LANGUAGE: ST
*)
IF F > 0.0 THEN
	tmp := 1000.0/F;
	CLK(PT := REAL_TO_TIME(tmp));
	Pulse(in := clk.Q, pt := REAL_TO_TIME(tmp*DC));
	Q := pulse.Q;
END_IF;

(* revision history

hm	25. feb 2007	rev 1.1
	recoded in st for better performance and better portability

hm	27. nov 2007	rev 1.2
	avoid divide by 0 when F = 0

hm	19. oct. 2008	rev 1.3
	changed type TP_R to TP_X because of name change
	improved performance

hm	11. mar. 2009	rev 1.4
	changed real constants to use dot syntax

*)
(*@KEY@: END_WORKSHEET *)
END_FUNCTION_BLOCK

(* ---- PWM_PW.ST ---- *)
(*@PROPERTIES_EX@
TYPE: POU
LOCALE: 0
IEC_LANGUAGE: ST
PLC_TYPE: independent
PROC_TYPE: independent
GROUP: ENGINEERING.SIGNAL_GENERATORS
*)
(*@KEY@:DESCRIPTION*)
version 1.5	11. mar. 2009
programmer 	oscat
tested BY	oscat

this signal generator generates a square wave signal which is specified by the frequency and the pulse width.

(*@KEY@:END_DESCRIPTION*)
FUNCTION_BLOCK PWM_PW

(*Group:Default*)

VAR_INPUT
	F :	REAL;
	PW :	TIME;
END_VAR

VAR_OUTPUT
	Q :	BOOL;
END_VAR

VAR
	clk :	CLK_Prg;
	pulse :	TP_X;
END_VAR

(*@KEY@: WORKSHEET
NAME: PWM_PW
IEC_LANGUAGE: ST
*)
IF F > 0.0 THEN
	CLK(PT := REAL_TO_TIME(1000.0 / F));
	Pulse(in := clk.Q, pt := pw);
	Q := pulse.Q;
END_IF;

(* revision history

hm	25. feb 2007	rev 1.1
	recoded in st for better performance and better portability

hm	27. nov 2007	rev 1.2
	avoid divide by 0 when F = 0

hm	9. dec 2007		rev 1.3
	corrected an error with F = 0

hm	19. oct. 2008	rev 1.4
	changed type tp_r to TP_x brecause of name change

hm	11. mar. 2009	rev 1.5
	changed real constants to use dot syntax

*)
(*@KEY@: END_WORKSHEET *)
END_FUNCTION_BLOCK

(* ---- RMP_B.ST ---- *)
(*@PROPERTIES_EX@
TYPE: POU
LOCALE: 0
IEC_LANGUAGE: ST
PLC_TYPE: independent
PROC_TYPE: independent
GROUP: ENGINEERING.SIGNAL_GENERATORS
*)
(*@KEY@:DESCRIPTION*)
version 2.0	23. oct. 2008
programmer 	oscat
tested BY	oscat

this ramp generator generates a byte wide ramp with 255 steps
the generator has an asynchronous set and reset
the ramp is controlled by PT which is the total ramp time for a full sweep from 0..255
an UD input controlls the direction Up or Down and the E input enables the ramp generation
a busy output indicates that the ramp is running, busy false means output is stable.
the outputs low and high will be true when the output has reached its max or min value.
(*@KEY@:END_DESCRIPTION*)
FUNCTION_BLOCK RMP_B

(*Group:Default*)

VAR_INPUT
	SET :	BOOL;
	PT :	TIME;
	E :	BOOL := TRUE;
	UP :	BOOL := TRUE;
	RST :	BOOL;
END_VAR

VAR_OUTPUT
	OUT :	BYTE;
	BUSY :	BOOL;
	HIGH :	BOOL;
	LOW :	BOOL;
END_VAR

VAR
	rmp :	_RMP_B;
END_VAR

(*@KEY@: WORKSHEET
NAME: RMP_B
IEC_LANGUAGE: ST
*)
(* generate ramp *)
rmp(dir := UP, E := E, TR := PT, RMP := out);
out := rmp.RMP;

(* set or reset operation *)
IF RST THEN
	out := BYTE#0;
ELSIF SET THEN
	out := BYTE#255;
END_IF;

(* checks for outputs stable and reset or set busy flag *)
low := out = BYTE#0;
high := out = BYTE#255;
busy := NOT (low OR high) AND E;

(* revision history

hm 5.10.2006	rev 1.1
	added busy output
hm 17.1.2007	rev 1.2
	renamed input ud to up for better usability
	deleted unused variable step

hm	17.9.2007		rev 1.3
	replaced time() with t_plc_ms() for compatibility reasons

hm	28. sep 2007	rev 1.4
	added outputs on and off
	busy is now disabled while en is false
	new coding for higher accuracy and performance

hm	5. oct 2007	rev 1.5
	added statements to allow for PT to be t#0s output jumps to max or min immediately

hm	25. dec 2007	rev 1.6
	improved code for better performance

hm	16. oct. 2008	rev 1.7
	improved code for better performance

hm	18. oct. 2008	rev 1.8
	added type conversion to avoid warnings
	changed input en to e for compatibility reasons

hm	23. oct. 2008	REV 	2.0
	new code using _RMP_B

*)
(*@KEY@: END_WORKSHEET *)
END_FUNCTION_BLOCK

(* ---- RMP_SOFT.ST ---- *)
(*@PROPERTIES_EX@
TYPE: POU
LOCALE: 0
IEC_LANGUAGE: ST
PLC_TYPE: independent
PROC_TYPE: independent
GROUP: ENGINEERING.SIGNAL_GENERATORS
*)
(*@KEY@:DESCRIPTION*)
version 2.0	26. oct. 2008
programmer 	oscat
tested BY	oscat

this soft on/off ramp generator generates a soft on and soft off ramp while the max on value is set by the input
the time for a full ramp can be set by config variables for up and down ramp.
(*@KEY@:END_DESCRIPTION*)
FUNCTION_BLOCK RMP_SOFT

(*Group:Default*)

VAR_INPUT
	IN :	BOOL;
	VAL :	BYTE;
	PT_ON :	TIME := T#100ms;
	PT_OFF :	TIME := T#100ms;
END_VAR

VAR_OUTPUT
	OUT :	BYTE := BYTE#00;
END_VAR

VAR
	rmp :	_RMP_B;
	tmp :	BYTE;
END_VAR

(*@KEY@: WORKSHEET
NAME: RMP_SOFT
IEC_LANGUAGE: ST
*)
tmp := SEL(in, BYTE#0, val);
IF tmp > out THEN
	(* we need to ramp down *)
	rmp(dir := TRUE, E := TRUE, TR := PT_ON, RMP := out);
	out := rmp.RMP;
	(* make sure out does not surpass tmp *)
	out := MIN(out, tmp);
ELSIF tmp < out THEN
	(* we need to ramp up *)
	rmp(dir := FALSE, E := TRUE, TR := PT_OFF, RMP := out);
	out := rmp.RMP;
	(* make sure out does not surpass tmp *)
	out := MAX(out, tmp);
ELSE
	(* no ramp necessary *)
	rmp(E := FALSE, RMP := out);
	out := rmp.RMP;
END_IF;

(* revision history

hm 22.1.2007	rev 1.1
	deleted unused variables X1 and I, X2 and X3

hm	17.9.2007	rev 1.2
	replaced time() with t_plc_ms() for compatibility reasons

hm	26. oct. 2008	2.0
	new code using _rmp_b
*)
(*@KEY@: END_WORKSHEET *)
END_FUNCTION_BLOCK

(* ---- RMP_W.ST ---- *)
(*@PROPERTIES_EX@
TYPE: POU
LOCALE: 0
IEC_LANGUAGE: ST
PLC_TYPE: independent
PROC_TYPE: independent
GROUP: ENGINEERING.SIGNAL_GENERATORS
*)
(*@KEY@:DESCRIPTION*)
version 2.0	23. oct. 2008
programmer 	oscat
tested BY	oscat

this ramp generator generates a Word wide ramp with 65535 steps
the generator has an asynchronous set and reset
the ramp is controlled by PT which is the total ramp time for a full sweep from 0..65535
an UD input controlls the direction Up or Down and the E input enables the ramp generation
a busy output indicates that the ramp is running, busy false means output is stable.
the outputs low and high will be true when the output has reached its max or min value.
(*@KEY@:END_DESCRIPTION*)
FUNCTION_BLOCK RMP_W

(*Group:Default*)

VAR_INPUT
	SET :	BOOL;
	PT :	TIME;
	E :	BOOL := TRUE;
	UP :	BOOL := TRUE;
	RST :	BOOL;
END_VAR

VAR_OUTPUT
	OUT :	WORD;
	BUSY :	BOOL;
	HIGH :	BOOL;
	LOW :	BOOL;
END_VAR

VAR
	rmp :	_RMP_W;
END_VAR

(*@KEY@: WORKSHEET
NAME: RMP_W
IEC_LANGUAGE: ST
*)
(* generate ramp *)
rmp(dir := UP, E := E, TR := PT, rmp := out);
out := rmp.RMP;

(* set or reset operation *)
IF RST THEN
	out := WORD#0;
ELSIF SET THEN
	out := WORD#65535;
END_IF;

(* checks for outputs stable and reset or set busy flag *)
low := out = WORD#0;
high := out = WORD#65535;
busy := NOT (low OR high) AND E;

(* revision history:

hm 4.10.2006		rev 1.1
	added the busy output which signals that the ramp is running.

hm 22.1.2007		rev 1.2
	deleted unused variable step

hm	17.9.2007		rev 1.3
	replaced time() with t_plc_ms() for compatibility reasons

hm	28. sep 2007	rev 1.4
	added outputs on and off
	busy is now disabled while en is false
	new coding for higher accuracy and performance

hm	5. oct 2007	rev 1.5
	added statements to allow for PT to be t#0s output jumps to max or min immediately

hm	2. dec 2007	rev 1.6
	corrected an error in calculation of step response

hm	25. dec 2007	rev 1.7
	corrected an error while step response was too slow for fast rise times

hm	16. oct. 2008	rev 1.8
	improved performance

hm	18. oct. 2008	rev 1.9
	renamed inout EN to E for compatibility reasons

hm	23. oct. 2008	rev 2.0
	new code using _RMP_W
*)
(*@KEY@: END_WORKSHEET *)
END_FUNCTION_BLOCK

(* ---- SCHEDULER.ST ---- *)
(*@PROPERTIES_EX@
TYPE: POU
LOCALE: 0
IEC_LANGUAGE: ST
PLC_TYPE: independent
PROC_TYPE: independent
GROUP: LOGIC.GENERATORS
*)
(*@KEY@:DESCRIPTION*)
version 1.0	28. sep 2008
programmer 	hugo
tested by	tobias

SCHEDULER is used to call programs or function blocks at specific intervals.
T0..T3 defines the interval times.
(*@KEY@:END_DESCRIPTION*)
FUNCTION_BLOCK SCHEDULER

(*Group:Default*)

VAR_INPUT
	E0 :	BOOL;
	E1 :	BOOL;
	E2 :	BOOL;
	E3 :	BOOL;
	T0 :	TIME;
	T1 :	TIME;
	T2 :	TIME;
	T3 :	TIME;
END_VAR

VAR_OUTPUT
	Q0 :	BOOL;
	Q1 :	BOOL;
	Q2 :	BOOL;
	Q3 :	BOOL;
END_VAR

VAR
	T_PLC_MS :	T_PLC_MS;
	init :	BOOL;
	s0 :	TIME;
	s1 :	TIME;
	s2 :	TIME;
	s3 :	TIME;
	tx :	TIME;
	c :	INT;
END_VAR

(*@KEY@: WORKSHEET
NAME: SCHEDULER
IEC_LANGUAGE: ST
*)
(* read sps timer *)
T_PLC_MS();
tx:= UDINT_TO_TIME(T_PLC_MS.T_PLC_MS);

IF NOT init THEN
	init := TRUE;
	s0 := tx - T0;
	s1 := tx - T1;
	s2 := tx - T2;
	s3 := tx - T3;
END_IF;

Q0 := FALSE;
Q1 := FALSE;
Q2 := FALSE;
Q3 := FALSE;

CASE c OF
	0: 	IF tx - s0 >= T0 THEN
			Q0 := E0;
			s0 := tx;
		END_IF;
		c := 1;
	1: 	IF tx - s1 >= T1 THEN
			Q1 := E1;
			s1 := tx;
		END_IF;
		c := 2;
	2: 	IF tx - s2 >= T2 THEN
			Q2 := E2;
			s2 := tx;
		END_IF;
		c := 3;
	3: 	IF tx - s3 >= T3 THEN
			Q3 := E3;
			s3 := tx;
		END_IF;
		c := 0;
END_CASE;

(* revision history

hm 28. sep. 2008		rev 1.0
	original version

*)
(*@KEY@: END_WORKSHEET *)
END_FUNCTION_BLOCK

(* ---- SCHEDULER_2.ST ---- *)
(*@PROPERTIES_EX@
TYPE: POU
LOCALE: 0
IEC_LANGUAGE: ST
PLC_TYPE: independent
PROC_TYPE: independent
GROUP: LOGIC.GENERATORS
*)
(*@KEY@:DESCRIPTION*)
version 1.0	29. sep 2008
programmer 	hugo
tested by	tobias

SCHEDULER_2 is used to call programs or function blocks at specific cycles.
C0..C3 defines after how many cycles the output becomes active.
O0..O3 defines a cycle offset at startup.
(*@KEY@:END_DESCRIPTION*)
FUNCTION_BLOCK SCHEDULER_2

(*Group:Default*)

VAR_INPUT
	E0 :	BOOL;
	E1 :	BOOL;
	E2 :	BOOL;
	E3 :	BOOL;
	C0 :	UINT;
	C1 :	UINT;
	C2 :	UINT;
	C3 :	UINT;
	O0 :	UINT;
	O1 :	UINT;
	O2 :	UINT;
	O3 :	UINT;
END_VAR

VAR_OUTPUT
	Q0 :	BOOL;
	Q1 :	BOOL;
	Q2 :	BOOL;
	Q3 :	BOOL;
END_VAR

VAR
	sx :	UINT;
END_VAR

(*@KEY@: WORKSHEET
NAME: SCHEDULER_2
IEC_LANGUAGE: ST
*)
Q0 := E0 AND (sx MOD C0 - O0 = UINT#0);
Q1 := E1 AND (sx MOD C1 - O1 = UINT#0);
Q2 := E2 AND (sx MOD C2 - O2 = UINT#0);
Q3 := E3 AND (sx MOD C3 - O3 = UINT#0);

(* increment cycle counter every cycle *)
sx := sx + UINT#1;

(* revision history
hm 29. sep. 2008		rev 1.0
	original version

*)
(*@KEY@: END_WORKSHEET *)
END_FUNCTION_BLOCK

(* ---- SEQUENCE_4.ST ---- *)
(*@PROPERTIES_EX@
TYPE: POU
LOCALE: 0
IEC_LANGUAGE: ST
PLC_TYPE: independent
PROC_TYPE: independent
GROUP: LOGIC.GENERATORS
*)
(*@KEY@:DESCRIPTION*)
version 1.4	17 sep 2007
programmer 	oscat
tested by	hans

sequence_4 enables run when a low to high transition is present on start.
a low to high transition on start will restart the sequencer at any time while a rst will hold the sequencer in reset while true.
after run is enabled with a rising edge on start the sequencer waits for wait0 on in0 to enable q0 which stays on for delay0.
the next cycle starts with wait1, continues with delay 1 and so on...
if an edge is not detected during the wait period, the sequencer will then display the error number on the status output.
the status numbers 1..4 are errors in step 0..3.
after the last step that sets q3, the sequencer leaves q3 on for delay3 and then resets to the initial state.
a step output will indicate the current step of the sequencer and will also be present with a fault condition.
after the first output is turened on the sequencer switches from q0 to q1 and so on, at any time there is only one output enabled.
if an input signal is not detected during a wait period, the sequencer will display the error number ( 1 for in0, 2 for in1 .... ).
when an error is present and the config variable stop_on_error is set then the sequencer will stop. otherwise it will continue.
The status output will also display 110 for waiting and 111 for sequence running.

(*@KEY@:END_DESCRIPTION*)
FUNCTION_BLOCK SEQUENCE_4

(*Group:Default*)

VAR_INPUT
	IN0 :	BOOL := TRUE;
	IN1 :	BOOL := TRUE;
	IN2 :	BOOL := TRUE;
	IN3 :	BOOL := TRUE;
	START :	BOOL;
	RST :	BOOL;
	WAIT0 :	TIME;
	DELAY0 :	TIME;
	WAIT1 :	TIME;
	DELAY1 :	TIME;
	WAIT2 :	TIME;
	DELAY2 :	TIME;
	WAIT3 :	TIME;
	DELAY3 :	TIME;
	STOP_ON_ERROR :	BOOL;
END_VAR

VAR_OUTPUT
	Q0 :	BOOL;
	Q1 :	BOOL;
	Q2 :	BOOL;
	Q3 :	BOOL;
	QX :	BOOL;
	RUN :	BOOL;
	STEP :	INT := -1;
	STATUS :	BYTE;
END_VAR

VAR
	last :	TIME;
	edge :	BOOL;
	tx :	TIME;
	init :	BOOL;
	T_PLC_MS :	T_PLC_MS;
END_VAR

(*@KEY@: WORKSHEET
NAME: SEQUENCE_4
IEC_LANGUAGE: ST
*)
(* read sps timer *)
T_PLC_MS();
tx:= UDINT_TO_TIME(T_PLC_MS.T_PLC_MS);

(* initialize on startup *)
IF NOT init THEN
	last := tx;
	init := TRUE;
	status := BYTE#110;
END_IF;

(* asynchronous reset *)
IF rst THEN
	step := -1;
	Q0 := FALSE;
	Q1 := FALSE;
	Q2 := FALSE;
	Q3 := FALSE;
	status := BYTE#110;
	run := FALSE;

(* edge on start input restarts the sequencer *)
ELSIF start AND NOT edge THEN
	step := 0;
	last := tx;
	status := BYTE#111;
	Q0 := FALSE;
	Q1 := FALSE;
	Q2 := FALSE;
	Q3 := FALSE;
	run := TRUE;
END_IF;
edge := start;

(* check if stop on status is necessary *)
IF status > BYTE#0 AND status < BYTE#100 AND stop_on_error THEN RETURN; END_IF;

(* sequence is running *)
IF run AND step = 0 THEN
	IF NOT q0 AND in0 AND tx - last <= wait0 THEN
		Q0 := TRUE;
		last := tx;
	ELSIF NOT q0 AND tx - last > wait0 THEN
		status := BYTE#1;
		run := FALSE;
	ELSIF q0 AND tx - last >= delay0 THEN
		step := 1;
		last := tx;
	END_IF;
END_IF;
IF run AND step = 1 THEN
	IF NOT q1 AND in1 AND tx - last <= wait1 THEN
		Q0 := FALSE;
		Q1 := TRUE;
		last := tx;
	ELSIF NOT q1 AND Tx - last > wait1 THEN
		status := BYTE#2;
		q0 := FALSE;
		run := FALSE;
	ELSIF q1 AND tx - last >= delay1 THEN
		step := 2;
		last := tx;
	END_IF;
END_IF;
IF run AND step = 2 THEN
	IF NOT q2 AND in2 AND tx - last <= wait2 THEN
		Q1 := FALSE;
		Q2 := TRUE;
		last := tx;
	ELSIF NOT q2 AND Tx - last > wait2 THEN
		status := BYTE#3;
		q1 := FALSE;
		run := FALSE;
	ELSIF q2 AND tx - last >= delay2 THEN
		step := 3;
		last := tx;
	END_IF;
END_IF;
IF run AND step = 3 THEN
	IF NOT q3 AND in3 AND tx - last <= wait3 THEN
		Q2 := FALSE;
		Q3 := TRUE;
		last := tx;
	ELSIF NOT q3 AND Tx - last > wait3 THEN
		status := BYTE#4;
		q2 := FALSE;
		run := FALSE;
	ELSIF q3 AND tx - last >= delay3 THEN
		step := -1;
		q3 := FALSE;
		run := FALSE;
		status := BYTE#110;
	END_IF;
END_IF;
QX := q0 OR q1 OR q2 OR q3;

(*
hm 1.10.06		rev 1.1
	corrected delay logic to be after event and not before
	added any output

hm 1.12.06		rev 1.2
	corrected failure in sequence logic.
	added init at startup to prevent from initial error after start.

hm 17.1.2007		rev 1.3
	changed output fault to status for better compatibility with other modules (ESR).
	added stop on error functionality and setup variable
	default for inputs in0..3 is true.
	renamed variable state to step

hm	17.sep 2007		rev 1.4
	replaced time() with T_PLC_MS() for compatibility reasons

*)
(*@KEY@: END_WORKSHEET *)
END_FUNCTION_BLOCK

(* ---- SEQUENCE_64.ST ---- *)
(*@PROPERTIES_EX@
TYPE: POU
LOCALE: 0
IEC_LANGUAGE: ST
PLC_TYPE: independent
PROC_TYPE: independent
GROUP: LOGIC.GENERATORS
*)
(*@KEY@:DESCRIPTION*)
version 1.0	29. jun. 2008
programmer 	hugo
tested by	oscat

sequence generates a sequence of states with a programmable length for each state.
(*@KEY@:END_DESCRIPTION*)
FUNCTION_BLOCK SEQUENCE_64

(*Group:Default*)

VAR_INPUT
	START :	BOOL;
	SMAX :	INT;
	RST :	BOOL;
END_VAR

VAR_OUTPUT
	STATE :	INT := INT#-1;
	TRIG :	BOOL;
END_VAR

VAR_IN_OUT
	PROG :	oscat_array64_time;
END_VAR

VAR
	T_PLC_MS :	T_PLC_MS;
	tx :	TIME;
	last :	TIME;
	edge :	BOOL;
END_VAR

(*@KEY@: WORKSHEET
NAME: SEQUENCE_64
IEC_LANGUAGE: ST
*)
(* read system timer *)
T_PLC_MS();
tx:= UDINT_TO_TIME(T_PLC_MS.T_PLC_MS);
TRIG := FALSE;

IF RST THEN
	STATE := -1;

(* start sequence *)
ELSIF START AND NOT edge THEN
	STATE := 0;
	last := tx;
	TRIG := TRUE;

(* sequence generator *)
ELSIF (STATE >= 0) THEN
	IF (tx - last) >= PROG[STATE] THEN
		STATE := INC2(STATE, 1, -1, SMAX);
		last := tx;
		TRIG := TRUE;
	END_IF;
END_IF;

edge := START;

(* revision history
hm	29. jun. 2008
	original version

*)
(*@KEY@: END_WORKSHEET *)
END_FUNCTION_BLOCK

(* ---- SEQUENCE_8.ST ---- *)
(*@PROPERTIES_EX@
TYPE: POU
LOCALE: 0
IEC_LANGUAGE: ST
PLC_TYPE: independent
PROC_TYPE: independent
GROUP: LOGIC.GENERATORS
*)
(*@KEY@:DESCRIPTION*)
version 1.4	17 sep 2007
programmer 	oscat
tested by		hans

sequence_8 enables run when a low to high transition is present on start.
a low to high transition on start will restart the sequencer at any time while a rst will hold the sequencer in reset while true.
after run is enabled with a rising edge on start the sequencer waits for wait0 on in0 to enable q0 which stays on for delay0.
the next cycle starts with wait1, continues with delay 1 and so on...
if an edge is not detected during the wait period, the sequencer will then display the error number on the status output.
The status numbers are 1 .. 8 for erros in step 0..7.
after the last step that sets q7, the sequencer leaves q7 on for delay7 and then resets to the initial state.
a step output will indicate the current step of the sequencer and will also be present with a fault condition.
after the first output is turened on the sequencer switches from q0 to q1 and so on, at any time there is only one output enabled.
if an input signal is not detected during a wait period, the sequencer will display the error number ( 1 for in0, 2 for in1 .... ).
when an error is present and the config variable stop_on_error is set then the sequencer will stop. otherwise it will continue.
The status output will also display 110 for waiting and 111 sequece running.
(*@KEY@:END_DESCRIPTION*)
FUNCTION_BLOCK SEQUENCE_8

(*Group:Default*)

VAR_INPUT
	IN0 :	BOOL := TRUE;
	IN1 :	BOOL := TRUE;
	IN2 :	BOOL := TRUE;
	IN3 :	BOOL := TRUE;
	IN4 :	BOOL := TRUE;
	IN5 :	BOOL := TRUE;
	IN6 :	BOOL := TRUE;
	IN7 :	BOOL := TRUE;
	START :	BOOL;
	RST :	BOOL;
	WAIT0 :	TIME;
	DELAY0 :	TIME;
	WAIT1 :	TIME;
	DELAY1 :	TIME;
	WAIT2 :	TIME;
	DELAY2 :	TIME;
	WAIT3 :	TIME;
	DELAY3 :	TIME;
	WAIT4 :	TIME;
	DELAY4 :	TIME;
	WAIT5 :	TIME;
	DELAY5 :	TIME;
	WAIT6 :	TIME;
	DELAY6 :	TIME;
	WAIT7 :	TIME;
	DELAY7 :	TIME;
	STOP_ON_ERROR :	BOOL;
END_VAR

VAR_OUTPUT
	Q0 :	BOOL;
	Q1 :	BOOL;
	Q2 :	BOOL;
	Q3 :	BOOL;
	Q4 :	BOOL;
	Q5 :	BOOL;
	Q6 :	BOOL;
	Q7 :	BOOL;
	QX :	BOOL;
	RUN :	BOOL;
	STEP :	INT := -1;
	STATUS :	BYTE;
END_VAR

VAR
	last :	TIME;
	edge :	BOOL;
	tx :	TIME;
	init :	BOOL;
	T_PLC_MS :	T_PLC_MS;
END_VAR

(*@KEY@: WORKSHEET
NAME: SEQUENCE_8
IEC_LANGUAGE: ST
*)
(* read sps timer *)
T_PLC_MS();
tx:= UDINT_TO_TIME(T_PLC_MS.T_PLC_MS);

(* initialize on startup *)
IF NOT init THEN
	last := tx;
	init := TRUE;
	status := BYTE#110;
END_IF;

(* asynchronous reset *)
IF rst THEN
	step := -1;
	Q0 := FALSE;
	Q1 := FALSE;
	Q2 := FALSE;
	Q3 := FALSE;
	Q4 := FALSE;
	Q5 := FALSE;
	Q6 := FALSE;
	Q7 := FALSE;
	status := BYTE#110;
	run := FALSE;

(* edge on start input restarts the sequencer *)
ELSIF start AND NOT edge THEN
	step := 0;
	last := tx;
	status := BYTE#111;
	Q0 := FALSE;
	Q1 := FALSE;
	Q2 := FALSE;
	Q3 := FALSE;
	Q4 := FALSE;
	Q5 := FALSE;
	Q6 := FALSE;
	Q7 := FALSE;
	run := TRUE;
END_IF;
edge := start;

(* check if stop on error is necessary *)
IF status > BYTE#0 AND status < BYTE#100 AND stop_on_error THEN RETURN; END_IF;

(* sequence is running *)
IF run AND step = 0 THEN
	IF NOT q0 AND in0 AND tx - last <= wait0 THEN
		Q0 := TRUE;
		last := tx;
	ELSIF NOT q0 AND tx - last > wait0 THEN
		status := BYTE#1;
		run := FALSE;
	ELSIF q0 AND tx - last >= delay0 THEN
		step := 1;
		last := tx;
	END_IF;
END_IF;
IF run AND step = 1 THEN
	IF NOT q1 AND in1 AND tx - last <= wait1 THEN
		Q0 := FALSE;
		Q1 := TRUE;
		last := tx;
	ELSIF NOT q1 AND Tx - last > wait1 THEN
		status := BYTE#2;
		q0 := FALSE;
		run := FALSE;
	ELSIF q1 AND tx - last >= delay1 THEN
		step := 2;
		last := tx;
	END_IF;
END_IF;
IF run AND step = 2 THEN
	IF NOT q2 AND in2 AND tx - last <= wait2 THEN
		Q1 := FALSE;
		Q2 := TRUE;
		last := tx;
	ELSIF NOT q2 AND Tx - last > wait2 THEN
		status := BYTE#3;
		q1 := FALSE;
		run := FALSE;
	ELSIF q2 AND tx - last >= delay2 THEN
		step := 3;
		last := tx;
	END_IF;
END_IF;
IF run AND step = 3 THEN
	IF NOT q3 AND in3 AND tx - last <= wait3 THEN
		Q2 := FALSE;
		Q3 := TRUE;
		last := tx;
	ELSIF NOT q3 AND Tx - last > wait3 THEN
		status := BYTE#4;
		q2 := FALSE;
		run := FALSE;
	ELSIF q3 AND tx - last >= delay3 THEN
		step := 4;
		last := tx;
	END_IF;
END_IF;
IF run AND step = 4 THEN
	IF NOT q4 AND in4 AND tx - last <= wait4 THEN
		Q3 := FALSE;
		Q4 := TRUE;
		last := tx;
	ELSIF NOT q4 AND Tx - last > wait4 THEN
		status := BYTE#5;
		q3 := FALSE;
		run := FALSE;
	ELSIF q4 AND tx - last >= delay4 THEN
		step := 5;
		last := tx;
	END_IF;
END_IF;
IF run AND step = 5 THEN
	IF NOT q5 AND in5 AND tx - last <= wait5 THEN
		Q4 := FALSE;
		Q5 := TRUE;
		last := tx;
	ELSIF NOT q5 AND Tx - last > wait5 THEN
		status := BYTE#6;
		q4 := FALSE;
		run := FALSE;
	ELSIF q5 AND tx - last >= delay5 THEN
		step := 6;
		last := tx;
	END_IF;
END_IF;
IF run AND step = 6 THEN
	IF NOT q6 AND in6 AND tx - last <= wait6 THEN
		Q5 := FALSE;
		Q6 := TRUE;
		last := tx;
	ELSIF NOT q6 AND Tx - last > wait6 THEN
		status := BYTE#7;
		q5 := FALSE;
		run := FALSE;
	ELSIF q6 AND tx - last >= delay6 THEN
		step := 7;
		last := tx;
	END_IF;
END_IF;
IF run AND step = 7 THEN
	IF NOT q7 AND in7 AND tx - last <= wait7 THEN
		Q6 := FALSE;
		Q7 := TRUE;
		last := tx;
	ELSIF NOT q7 AND Tx - last > wait7 THEN
		status := BYTE#8;
		q6 := FALSE;
		run := FALSE;
	ELSIF q7 AND tx - last >= delay7 THEN
		step := -1;
		Q7 := FALSE;
		Run := FALSE;
		status := BYTE#110;
	END_IF;
END_IF;
QX := q0 OR q1 OR q2 OR q3 OR q4 OR q5 OR q6 OR q7;

(*
hm 1.10.06		rev 1.1
	corrected delay logic to be after event and not before
	added any output

hm 1.12.06		rev 1.2
	corrected failure in sequence logic.
	added init at startup to prevent from initial statuss after start.

hm 17.1.2007		rev 1.3
	changed output fault to status for better compatibility with other modules (ESR)
	added stop on error functionality and setup variable
	default for inputs in0..7 is true.
	renames variable state to step

hm	17.sep 2007		rev 1.4
	replaced time() with T_PLC_MS() for compatibility reasons

*)
(*@KEY@: END_WORKSHEET *)
END_FUNCTION_BLOCK

(* ---- SRAMP.ST ---- *)
(*@PROPERTIES_EX@
TYPE: POU
LOCALE: 0
IEC_LANGUAGE: ST
PLC_TYPE: independent
PROC_TYPE: independent
GROUP: ENGINEERING.AUTOMATION
*)
(*@KEY@:DESCRIPTION*)
version 1.1	11. mar. 2009
programmer 	hugo
tested by	tobias

RAMPS generates output signal which are slew rate and acceleration controlled.

(*@KEY@:END_DESCRIPTION*)
FUNCTION_BLOCK SRAMP

(*Group:Default*)

VAR_INPUT
	X :	REAL;
	A_UP :	REAL;
	A_DN :	REAL;
	VU_MAX :	REAL;
	VD_MAX :	REAL;
	LIMIT_HIGH :	REAL;
	LIMIT_LOW :	REAL;
	RST :	BOOL;
END_VAR

VAR_OUTPUT
	Y :	REAL;
	V :	REAL;
END_VAR

VAR
	cycle_time :	TC_S;
	init :	BOOL;
END_VAR

(*@KEY@: WORKSHEET
NAME: SRAMP
IEC_LANGUAGE: ST
*)
(* read the system_time in microseconds *)
cycle_time();

(* assure range of inputs *)
A_up := MAX(0.0,A_UP);
A_dn := MIN(0.0,A_dn);
VU_max := MAX(0.0,VU_max);
VD_max := MIN(0.0,VD_MAX);

(* calculate the output offset *)
IF rst OR NOT init THEN
	init := TRUE;
	Y := 0.0;
	V := 0.0;
ELSIF X = Y THEN
	v := 0.0;
ELSIF X > Y THEN
	(* output is too low >> ramp up and brake at the end *)
	(* accelerate the speed and limit to vu_max *)
	v := MIN(v + A_UP * cycle_time.TC, vu_max);
	(* calculate the max speed to be able to brake and select the lowest *)
	v := MIN(SQRT((Y-X) * 2.0 * A_DN), v);
	(* calculate the output and obey limits *)
	y := LIMIT(limit_low, y + MIN(v * cycle_time.TC, X-Y), limit_high);
ELSIF X < Y THEN
	(* output is too high >> ramp dn and brake at the end *)
	(* accelerate the speed and limit to vd_max *)
	v := MAX(v + A_DN * cycle_time.TC, vd_max);
	(* calculate the max speed to be able to brake and select the lowest *)
	v := MAX(-SQRT((Y-X) * 2.0 * A_UP), v);
	(* calculate the output and obey limits *)
	y := LIMIT(limit_low, y + MAX(v * cycle_time.TC, X-Y), limit_high);
END_IF;

(* revision history
hm	13. mar. 2008	rev 1.0
	original version

hm	11. mar. 2009	rev 1.1
	real constants updated to new systax using dot

*)

(*@KEY@: END_WORKSHEET *)
END_FUNCTION_BLOCK

(* ---- STACK_16.ST ---- *)
(*@PROPERTIES_EX@
TYPE: POU
LOCALE: 0
IEC_LANGUAGE: ST
PLC_TYPE: independent
PROC_TYPE: independent
GROUP: LOGIC.MEMORY
*)
(*@KEY@:DESCRIPTION*)
version 2.0	25. jul 2009
programmer 	hugo
tested by	oscat

16 Dword STACK memory

(*@KEY@:END_DESCRIPTION*)
FUNCTION_BLOCK STACK_16

(*Group:Default*)

VAR_INPUT
	DIN :	DWORD;
	E :	BOOL := TRUE;
	RD :	BOOL;
	WD :	BOOL;
	RST :	BOOL;
END_VAR

VAR_OUTPUT
	DOUT :	DWORD;
	EMPTY :	BOOL := TRUE;
	FULL :	BOOL;
END_VAR

VAR
	pt :	INT;
	stack :	oscat_ardw_0_15;
END_VAR

(*@KEY@: WORKSHEET
NAME: STACK_16
IEC_LANGUAGE: ST
*)
IF RST THEN
	(* asynchronous reset for the fifo *)
	pt := 0;
	EMPTY := TRUE;
	FULL := FALSE;
	Dout := DWORD#0;
ELSIF E THEN
	IF NOT EMPTY AND RD THEN
		(* read one element *)
		pt := pt - 1;
		Dout := stack[pt];
		EMPTY := pt = 0;
		FULL := FALSE;
	END_IF;
	IF NOT FULL AND WD THEN
		(* write one element *)
		stack[pt] := Din;
		pt := pt + 1;
		FULL := pt > 15;
		EMPTY := FALSE;
	END_IF;
END_IF;

(* revision history
hm	4. aug. 2006	rev 1.0
	original version

hm	19. feb 2008	rev 1.1
	performance improvements

hm	17. oct. 2008	rev 1.2
	deleted unnecessary init with 0

hm	27. oct. 2008	rev 1.3
	optimized performance

hm	25. jul 2009	rev 2.0
	changed inputs to allow simultsaneous read and write
*)

(*@KEY@: END_WORKSHEET *)
END_FUNCTION_BLOCK

(* ---- STACK_32.ST ---- *)
(*@PROPERTIES_EX@
TYPE: POU
LOCALE: 0
IEC_LANGUAGE: ST
PLC_TYPE: independent
PROC_TYPE: independent
GROUP: LOGIC.MEMORY
*)
(*@KEY@:DESCRIPTION*)
version 2.0	25. jul 2009
programmer 	hugo
tested by	oscat

32 Dword STACK memory
(*@KEY@:END_DESCRIPTION*)
FUNCTION_BLOCK STACK_32

(*Group:Default*)

VAR_INPUT
	DIN :	DWORD;
	E :	BOOL := TRUE;
	RD :	BOOL;
	WD :	BOOL;
	RST :	BOOL;
END_VAR

VAR_OUTPUT
	DOUT :	DWORD;
	EMPTY :	BOOL := TRUE;
	FULL :	BOOL;
END_VAR

VAR
	pt :	INT;
	stack :	oscat_ardw_0_31;
END_VAR

(*@KEY@: WORKSHEET
NAME: STACK_32
IEC_LANGUAGE: ST
*)
IF RST THEN
	(* asynchronous reset for the fifo *)
	pt := 0;
	EMPTY := TRUE;
	FULL := FALSE;
	Dout := DWORD#0;
ELSIF E THEN
	IF NOT EMPTY AND RD THEN
		(* read one element *)
		pt := pt - 1;
		Dout := stack[pt];
		EMPTY := pt = 0;
		FULL := FALSE;
	END_IF;
	IF NOT FULL AND WD THEN
		(* write one element *)
		stack[pt] := Din;
		pt := pt + 1;
		FULL := pt > 31;
		EMPTY := FALSE;
	END_IF;
END_IF;

(* revision history
hm	4. aug. 2006	rev 1.0
	original version

hm	19. feb 2008	rev 1.1
	performance improvements

hm	17. oct. 2008	rev 1.2
	deleted unnecessary init with 0

ks	27. oct. 2008	rev 1.3
	optimized performance

hm	25. jul 2009	rev 2.0
	changed inputs to allow simultsaneous read and write

*)

(*@KEY@: END_WORKSHEET *)
END_FUNCTION_BLOCK

(* ---- STAIR2.ST ---- *)
(*@PROPERTIES_EX@
TYPE: POU
LOCALE: 0
IEC_LANGUAGE: ST
PLC_TYPE: independent
PROC_TYPE: independent
GROUP: ENGINEERING.SIGNAL_PROCESSING
*)
(*@KEY@:DESCRIPTION*)
version 1.4	10. mar. 2009
programmer 	hugo
tested by	oscat

the function stair2 converts an anlog input signal to a staircase like output.
D is the step width for the output signal. the output will use D as a hysteresis for a stairchange.
if D = 0 then the output follows the input without a chage.
(*@KEY@:END_DESCRIPTION*)
FUNCTION_BLOCK STAIR2

(*Group:Default*)

VAR_INPUT
	X :	REAL;
	D :	REAL;
END_VAR

VAR_OUTPUT
	Y :	REAL;
END_VAR

(*@KEY@: WORKSHEET
NAME: STAIR2
IEC_LANGUAGE: ST
*)
IF D > 0.0 THEN
	IF X >= Y + D OR X <= Y - D THEN Y := INT_TO_REAL(FLOOR(X/D)) * D; END_IF;
ELSE
	Y := X;
END_IF;

(* revision history
hm	28 jan 2007		rev 1.0
	original version

hm	27. dec 2007	rev 1.1
	changed code for better performance

hm	30. jun. 2008	rev 1.2
	added type conversions to avoid warnings under codesys 3.0

ks	26. oct. 2008	rev 1.3
	improved code

hm	10. mar. 2009	rev 1.4
	real constants updated to new systax using dot

*)
(*@KEY@: END_WORKSHEET *)
END_FUNCTION_BLOCK

(* ---- TICKER.ST ---- *)
(*@PROPERTIES_EX@
TYPE: POU
LOCALE: 0
IEC_LANGUAGE: ST
PLC_TYPE: independent
PROC_TYPE: independent
GROUP: STRINGS
*)
(*@KEY@:DESCRIPTION*)
version 1.2	29. mar. 2008
programmer 	hugo
tested by	tobias

Ticker sends a substring of text with length N every TD Milliseconds to generate a ticker.
(*@KEY@:END_DESCRIPTION*)
FUNCTION_BLOCK TICKER

(*Group:Default*)

VAR_INPUT
	N :	INT;
	PT :	TIME;
	TEXT :	STRING;
END_VAR

VAR_OUTPUT
	DISPLAY :	STRING;
END_VAR

VAR
	delay :	TP;
	rollout :	STRING;
	text_len :	INT;
	rollout_step :	INT;
	step :	INT;
END_VAR

(*@KEY@: WORKSHEET
NAME: TICKER
IEC_LANGUAGE: ST
*)
(* generate next ticker when delay is low *)
text_len := LEN(text);

IF N < text_len THEN
	IF NOT delay.Q THEN

		IF step > text_len THEN
            rollout_step := 0;
            rollout := '';
            step := 0;
        END_IF;

        IF step + N > text_len THEN
		    (* increase step for next tick *)
		    step := step + 1;
            rollout_step := rollout_step +1;
		    (* extract dispay from text *)
		    display := MID(text, N - rollout_step, step);
            rollout := CONCAT(rollout,'#');
            display := CONCAT(display,rollout);
        ELSE
		    (* increase step for next tick *)
		    step := step + 1;
		    (* extract dispay from text *)
		    display := MID(text, N, step);
        END_IF;

		(* set delay timer for next tick *)
		delay(in := TRUE, PT := PT);
	ELSE;
		(* execute delay timer *)
		delay(in := FALSE);
	END_IF;
ELSE
	display := text;
END_IF;

(* revision history
hm	4. dec. 2007	rev 1.0
	original version

hm	15. dec. 2007	rev 1.1
	step now starts at 1 instaed of 0

hm	29. mar. 2008	rev 1.2
	changed STRING to STRING(STRING_LENGTH)
*)
(*@KEY@: END_WORKSHEET *)
END_FUNCTION_BLOCK

(* ---- TOF_1.ST ---- *)
(*@PROPERTIES_EX@
TYPE: POU
LOCALE: 0
IEC_LANGUAGE: ST
PLC_TYPE: independent
PROC_TYPE: independent
GROUP: LOGIC.GENERATORS
*)
(*@KEY@:DESCRIPTION*)
version 1.0	17. jul. 2008
programmer 	hugo
tested by	oscat

TOF_1 will extend a pulse on input in for PT seconds.
in addition the timer can be cleared asynchronously with rst.
TOF_1 is the same function as TOF from the standard LIB except the asynchronous reset input.
(*@KEY@:END_DESCRIPTION*)
FUNCTION_BLOCK TOF_1

(*Group:Default*)

VAR_INPUT
	IN :	BOOL;
	PT :	TIME;
	RST :	BOOL;
END_VAR

VAR_OUTPUT
	Q :	BOOL;
END_VAR

VAR
	start :	TIME;
	tx :	TIME;
	T_PLC_MS :	T_PLC_MS;
END_VAR

(*@KEY@: WORKSHEET
NAME: TOF_1
IEC_LANGUAGE: ST
*)
(* read system timer *)
T_PLC_MS();
tx:= UDINT_TO_TIME(T_PLC_MS.T_PLC_MS);

IF RST THEN
	Q := FALSE;
ELSIF IN THEN
	Q := TRUE;
	start := tx;
ELSIF tx - start >= PT THEN
	Q := FALSE;
END_IF;

(* revision history
hm	17. jul. 2008	rev 1.0
	original version

*)
(*@KEY@: END_WORKSHEET *)
END_FUNCTION_BLOCK

(* ---- TONOF.ST ---- *)
(*@PROPERTIES_EX@
TYPE: POU
LOCALE: 0
IEC_LANGUAGE: ST
PLC_TYPE: independent
PROC_TYPE: independent
GROUP: LOGIC.GENERATORS
*)
(*@KEY@:DESCRIPTION*)
version 1.2	21. jul 2009
programmer 	hugo
tested by	tobias

TONOF generated a TON and TOF Delay for the Input N TON (T1) and TOF (T2) can be configured separately

(*@KEY@:END_DESCRIPTION*)
FUNCTION_BLOCK TONOF

(*Group:Default*)

VAR_INPUT
	IN :	BOOL;
	T_ON :	TIME;
	T_OFF :	TIME;
END_VAR

VAR_OUTPUT
	Q :	BOOL;
END_VAR

VAR
	X :	TON;
	old :	BOOL;
	mode :	BOOL;
END_VAR

(*@KEY@: WORKSHEET
NAME: TONOF
IEC_LANGUAGE: ST
*)
IF IN XOR old THEN
  X(IN := FALSE, PT := SEL_TIME(IN,T_OFF,T_ON));
  mode := IN;
  old := IN;
END_IF;
X(IN := TRUE);
IF X.Q THEN Q := mode;END_IF;

(* revision history
hm	10. dec 2007	rev 1.0
	original version

hm	17. sep. 2007	rev 1.1
	improved performance

hm	21. jul. 2009	rev 1.2
	fixed a timing probelm

*)

(*@KEY@: END_WORKSHEET *)
END_FUNCTION_BLOCK

(* ---- TP_1.ST ---- *)
(*@PROPERTIES_EX@
TYPE: POU
LOCALE: 0
IEC_LANGUAGE: ST
PLC_TYPE: independent
PROC_TYPE: independent
GROUP: LOGIC.GENERATORS
*)
(*@KEY@:DESCRIPTION*)
version 1.0	28. jun. 2008
programmer 	hugo
tested by	oscat

TP_1 generates a pulse every time it is calles with in := TRUE.
in addition the timer can be cleared asynchronously with rst.
the timer can be retriggered as often as necessary. it will count PT from the last trigger.
(*@KEY@:END_DESCRIPTION*)
FUNCTION_BLOCK TP_1

(*Group:Default*)

VAR_INPUT
	IN :	BOOL;
	PT :	TIME;
	RST :	BOOL;
END_VAR

VAR_OUTPUT
	Q :	BOOL;
END_VAR

VAR
	tx :	TIME;
	start :	TIME;
	ix :	BOOL;
	T_PLC_MS :	T_PLC_MS;
END_VAR

(*@KEY@: WORKSHEET
NAME: TP_1
IEC_LANGUAGE: ST
*)
(* read system timer *)
(* read system_time *)
T_PLC_MS();
tx := UDINT_TO_TIME(T_PLC_MS.T_PLC_MS);

IF RST THEN
	Q := FALSE;
ELSIF IN AND NOT ix THEN
	Q := TRUE;
	start := tx;
ELSIF tx - start >= PT THEN
	Q := FALSE;
END_IF;

ix:= IN;

(* revision history
hm	28. jun. 2008
	original version

*)
(*@KEY@: END_WORKSHEET *)
END_FUNCTION_BLOCK

(* ---- TP_1D.ST ---- *)
(*@PROPERTIES_EX@
TYPE: POU
LOCALE: 0
IEC_LANGUAGE: ST
PLC_TYPE: independent
PROC_TYPE: independent
GROUP: LOGIC.GENERATORS
*)
(*@KEY@:DESCRIPTION*)
version 1.0	28. jun. 2008
programmer 	hugo
tested by	oscat

TP_2 generates a pulse every time it is calles with in := TRUE.
the module will reset IN by itself so no clearing of in is necessary.
in addition the timer can be cleared asynchronously with rst.
also the rst input is cleared by the module itself.
the timer can be retriggered as often as necessary. it will count PT from the last trigger.
after the time PT1 is elapsed, the timer blocks itself for PT2 and only allow new sequences after PT2 has elapsed.
(*@KEY@:END_DESCRIPTION*)
FUNCTION_BLOCK TP_1D

(*Group:Default*)

VAR_INPUT
	IN :	BOOL;
	PT1 :	TIME;
	PTD :	TIME;
	RST :	BOOL;
END_VAR

VAR_OUTPUT
	Q :	BOOL;
	W :	BOOL;
END_VAR

VAR
	tx :	TIME;
	start :	TIME;
	ix :	BOOL;
	T_PLC_MS :	T_PLC_MS;
END_VAR

(*@KEY@: WORKSHEET
NAME: TP_1D
IEC_LANGUAGE: ST
*)
(* read system_time *)
T_PLC_MS();
tx := UDINT_TO_TIME(T_PLC_MS.T_PLC_MS);

IF RST THEN
	Q := FALSE;
	rst := FALSE;
	W := FALSE;
ELSIF W THEN
	IF tx - start >= PTD THEN
		W := FALSE;
	END_IF;
ELSIF IN AND NOT ix THEN
	Q := TRUE;
	start := tx;
	in := FALSE;
ELSIF tx - start >= PT1 THEN
	Q := FALSE;
	W := TRUE;
	start := tx;
END_IF;

ix := IN;

(* revision history
hm	28. jun. 2008
	original version

*)
(*@KEY@: END_WORKSHEET *)
END_FUNCTION_BLOCK

(* ---- TP_X.ST ---- *)
(*@PROPERTIES_EX@
TYPE: POU
LOCALE: 0
IEC_LANGUAGE: ST
PLC_TYPE: independent
PROC_TYPE: independent
GROUP: LOGIC.GENERATORS
*)
(*@KEY@:DESCRIPTION*)
version 1.3	17. dec. 2008
programmer 	hugo
tested by	oscat

retriggerable edge triggered pulse similar to TP but with a retrigger function
if the pt input is 0 then output is always low.
(*@KEY@:END_DESCRIPTION*)
FUNCTION_BLOCK TP_X

(*Group:Default*)

VAR_INPUT
	IN :	BOOL;
	PT :	TIME;
END_VAR

VAR_OUTPUT
	Q :	BOOL;
	ET :	TIME;
END_VAR

VAR
	edge :	BOOL;
	start :	TIME;
	tx :	TIME;
	T_PLC_MS :	T_PLC_MS;
END_VAR

(*@KEY@: WORKSHEET
NAME: TP_X
IEC_LANGUAGE: ST
*)
(* read system_time *)
T_PLC_MS();
tx := UDINT_TO_TIME(T_PLC_MS.T_PLC_MS);

(* rising edge trigger *)
IF IN AND NOT edge THEN
	start := tx;
	Q := PT > t#0ms;
ELSIF Q THEN
	ET := tx - start;
	IF ET >= PT THEN
		Q := FALSE;
		ET := t#0ms;
	END_IF;
END_IF;
edge := IN;

(* revision history
hm	4. aug 2006		rev 1.0
	original version

hm	17. sep 2007	rev 1.1
	replaced time() with T_PLC_MS() for compatibility reasons

hm	19. oct. 2008	rev 1.2
	renamed to TP_R to TP_X for compatibility reasons

hm	17. dec. 2008	rev 1.3
	code optimized

*)
(*@KEY@: END_WORKSHEET *)
END_FUNCTION_BLOCK

(* ---- TUNE.ST ---- *)
(*@PROPERTIES_EX@
TYPE: POU
LOCALE: 0
IEC_LANGUAGE: ST
PLC_TYPE: independent
PROC_TYPE: independent
GROUP: ENGINEERING.AUTOMATION
*)
(*@KEY@:DESCRIPTION*)
version 1.2	11. mar. 2009
programmer 	hugo
tested by	tobias

tune generates an output signal which is set by input switches.
up to 4 switsches can be used to tune the signal up or down.

(*@KEY@:END_DESCRIPTION*)
FUNCTION_BLOCK TUNE

(*Group:Default*)

VAR_INPUT
	SET :	BOOL;
	SU :	BOOL;
	SD :	BOOL;
	RST :	BOOL;
	SS :	REAL := 0.1;
	LIMIT_L :	REAL;
	LIMIT_H :	REAL := 100.0;
	RST_VAL :	REAL;
	SET_VAL :	REAL := 100.0;
	T1 :	TIME := T#500ms;
	T2 :	TIME := T#2s;
	S1 :	REAL := 2.0;
	S2 :	REAL := 10.0;
END_VAR

VAR_OUTPUT
	Y :	REAL;
END_VAR

VAR
	tx :	UDINT;
	start :	UDINT;
	start2 :	UDINT;
	state :	INT;
	in :	BOOL;
	step :	REAL;
	speed :	REAL;
	Y_start :	REAL;
	Y_start2 :	REAL;
	T_PLC_MS :	T_PLC_MS;
END_VAR

(*@KEY@: WORKSHEET
NAME: TUNE
IEC_LANGUAGE: ST
*)
(* read system_time *)
T_PLC_MS();
tx:= T_PLC_MS.T_PLC_MS;

IF rst THEN
	Y := RST_val;
	state := 0;
ELSIF set THEN
	Y := SET_val;
	state := 0;
ELSIF state > 0 THEN
	(* key has been pushed state machine operating *)
	(* first read the correct input *)
	IF state = 1 THEN
		(* step up *)
		in := su;
	ELSE
		(* step down *)
		in := sd;
	END_IF;
	(* check for single step operation *)
	IF NOT in AND tx - start <= TIME_TO_UDINT(T1) THEN
		Y := Y_start + step;
		state := 0;
	(* check if fast ramp needs to be generated *)
	ELSIF in AND tx - start >= TIME_TO_UDINT(T2) THEN
		Y := Y_start2 + UDINT_TO_REAL(tx - start2) * s2 / speed;
	(* check if slow ramp needs to be generated *)
	ELSIF in AND tx - start >= TIME_TO_UDINT(T1) THEN
		Y := Y_start + UDINT_TO_REAL(tx - start - TIME_TO_UDINT(T1)) * S1 / speed;
		start2 := tx;
		Y_start2 := Y;
	ELSIF NOT in THEN
		state := 0;
	END_IF;
ELSIF su THEN
	(* slow step up *)
	state := 1;
	start := tx;
	step := ss;
	speed := 1000.0;
	Y_start := Y;
ELSIF sd THEN
	(* slow step down *)
	state := 2;
	start := tx;
	step := -ss;
	speed := -1000.0;
	Y_start := Y;
END_IF;

(* make sure output does not exceed limits *)
Y := LIMIT(LIMIT_L, Y, LIMIT_H);

(* revision history
hm	3.11.2007		rev 1.0
	original version

hm	16. mar. 2008	rev 1.1
	added type conversions to avoid warnings under codesys 3.0

hm	11. mar. 2009	rev 1.2
	real constants updated to new systax using dot

*)
(*@KEY@: END_WORKSHEET *)
END_FUNCTION_BLOCK

(* ---- TUNE2.ST ---- *)
(*@PROPERTIES_EX@
TYPE: POU
LOCALE: 0
IEC_LANGUAGE: ST
PLC_TYPE: independent
PROC_TYPE: independent
GROUP: ENGINEERING.AUTOMATION
*)
(*@KEY@:DESCRIPTION*)
version 1.2	11. mar. 2009
programmer 	hugo
tested by	tobias

tune2 generates an output signal which is set by input switches.
up to 4 switsches can be used to tune the signal up or down.

(*@KEY@:END_DESCRIPTION*)
FUNCTION_BLOCK TUNE2

(*Group:Default*)

VAR_INPUT
	SET :	BOOL;
	SU :	BOOL;
	SD :	BOOL;
	FU :	BOOL;
	FD :	BOOL;
	RST :	BOOL;
	SS :	REAL := 0.1;
	FS :	REAL := 5.0;
	LIMIT_L :	REAL;
	LIMIT_H :	REAL := 100.0;
	RST_VAL :	REAL;
	SET_VAL :	REAL := 100.0;
	TR :	TIME := T#500ms;
	S1 :	REAL := 2.0;
	S2 :	REAL := 10.0;
END_VAR

VAR_OUTPUT
	Y :	REAL;
END_VAR

VAR
	tx :	UDINT;
	start :	UDINT;
	state :	INT;
	in :	BOOL;
	step :	REAL;
	speed :	REAL;
	Y_start :	REAL;
	T_PLC_MS :	T_PLC_MS;
END_VAR

(*@KEY@: WORKSHEET
NAME: TUNE2
IEC_LANGUAGE: ST
*)
(* read system time *)
T_PLC_MS();
tx:= T_PLC_MS.T_PLC_MS;

IF rst THEN
	Y := RST_val;
	state := 0;
ELSIF set THEN
	Y := SET_val;
	state := 0;
ELSIF state > 0 THEN
	(* key has been pushed state machine operating *)
	(* first read the correct input *)
	CASE state OF
		1 :	(* slow up *)
			in := su;
		2 :	(* slow down *)
			in := sd;
		3 :	(* fast up *)
			in := fu;
		4 :	(* fast down *)
			in := fd;
	END_CASE;
	(* check for single step operation *)
	IF NOT in AND tx - start <= TIME_TO_UDINT(TR) THEN
		Y := Y_start + step;
		state := 0;
	(* check if ramp needs to be generated *)
	ELSIF in AND tx - start >= TIME_TO_UDINT(TR) THEN
		Y := Y_start + UDINT_TO_REAL(tx - start - TIME_TO_UDINT(TR)) * speed;
	ELSIF NOT in THEN
		state := 0;
	END_IF;
ELSIF su THEN
	(* slow step up *)
	state := 1;
	start := tx;
	step := ss;
	speed := s1 * 1.0E-3;
	Y_start := Y;
ELSIF sd THEN
	(* slow step down *)
	state := 2;
	start := tx;
	step := -ss;
	speed := -s1 * 1.0E-3;
	Y_start := Y;
ELSIF fu THEN
	(* fast step up *)
	state := 3;
	start := tx;
	step := fs;
	speed := s2 * 1.0E-3;
	y_start := Y;
ELSIF fd THEN
	(* fast step down *)
	state := 4;
	start := tx;
	step := -fs;
	speed := -s2 * 1.0E-3;
	y_start := Y;
END_IF;

(* make sure output does not exceed limits *)
Y := LIMIT(LIMIT_L, Y, LIMIT_H);

(* revision history
hm	3.11.2007		rev 1.0
	original version

hm	16. 3. 2008	rev 1.1
	added type conversions to avoid warnings in codesys 3.0
	improved performance

hm	11. mar. 2009	rev 1.2
	real constants updated to new systax using dot

*)
(*@KEY@: END_WORKSHEET *)
END_FUNCTION_BLOCK

(* ---- AIN.ST ---- *)
(*@PROPERTIES_EX@
TYPE: POU
LOCALE: 0
IEC_LANGUAGE: ST
PLC_TYPE: independent
PROC_TYPE: independent
GROUP: ENGINEERING.SIGNAL_PROCESSING
*)
(*@KEY@:DESCRIPTION*)
version 1.5	16 mar 2008
programmer 	oscat
tested by	tobias

Ain converts signals from A/D converters or other digital sources to an internal real value
the lowest number of bits are extracted from the input word and the sign will be extracted if available separately.
the output signal is then conditioned to range from low to high values for a 0 to max value on the analog inputs:
for example a 15bit input (bits := 12) with sign at bit 15 (0..15) will deliver 0.0 (low value at 0) for an input value of 2#0000_0000_0000
an input value of 2#1111_1111_1111 will deliver 10.0 on the output (high value set to 10).
(*@KEY@:END_DESCRIPTION*)
FUNCTION AIN:REAL

(*Group:Default*)

VAR_INPUT
	IN :	DWORD;
	BITS :	BYTE;
	SIGN :	BYTE;
	LOW :	REAL;
	HIGH :	REAL;
END_VAR

VAR
	temp1 :	DWORD;
	temp2 :	DWORD;
	sx :	BOOL;
END_VAR

(*@KEY@: WORKSHEET
NAME: AIN
IEC_LANGUAGE: ST
*)
(* extract the sign bit *)
IF sign < BYTE#32 THEN
	temp1 := SHR_DWORD(in, _BYTE_TO_INT(sign));
	sx := BIT_OF_DWORD(temp1,0); (* temp1.X0 *)
ELSE
	sx := FALSE;
END_IF;
temp1 := SHR_DWORD(DWORD#16#FFFFFFFF,32 - _BYTE_TO_INT(bits));
temp2 := in AND temp1;
AIN := (high - low)* _DWORD_TO_REAL(temp2) / _DWORD_TO_REAL(temp1) + low;
IF sx THEN AIN := -AIN; END_IF;

(* revision history
hm 18.8.2006	rev 1.1
	fixed an error with low value negative and high value 0.

hm 19.1.2007	rev 1.2
	fixed an error with sign bit.

hm	13.9.2007	rev 1.3
	changed code to avoid warning under codesys 2.8.1

hm	2. dec 2007	rev 1.4
	changed code for better performance

hm	16. mar 2008	rev 1.5
	added type conversions to avoid warnings under codesys 30
*)
(*@KEY@: END_WORKSHEET *)
END_FUNCTION

(* ---- AOUT.ST ---- *)
(*@PROPERTIES_EX@
TYPE: POU
LOCALE: 0
IEC_LANGUAGE: ST
PLC_TYPE: independent
PROC_TYPE: independent
GROUP: ENGINEERING.SIGNAL_PROCESSING
*)
(*@KEY@:DESCRIPTION*)
version 1.4	23 feb 2008
programmer 	oscat
tested by	tobias

this module conditions an internal real value for D/A converter.
Aout converts and internal real value to a word for an D/A converter or other output devices.
The input value is converted to a n-bit wide output and a sign bit is set separately as specified.
the outout min value is set for the specified min input value and the max output is set for the max input value.
an input higher or lower then the max or min value will set the respective max or min value or the output.
in value or the output.
(*@KEY@:END_DESCRIPTION*)
FUNCTION AOUT:DWORD

(*Group:Default*)

VAR_INPUT
	IN :	REAL;
	BITS :	BYTE;
	SIGN :	BYTE;
	LOW :	REAL;
	HIGH :	REAL;
END_VAR

VAR
	in2 :	REAL;
	sx :	BOOL;
END_VAR

(*@KEY@: WORKSHEET
NAME: AOUT
IEC_LANGUAGE: ST
*)
(* if sign bit is defined *)
IF sign < BYTE#32 THEN
	sx := sign_R(in);
	in2 := ABS(in);
ELSE
	in2 := in;
END_IF;

(* begrenze in auf die zulässigen werte *)
in2 := LIMIT(low, in2, high);

(* Berechne den Ausgangswert *)
Aout := _REAL_TO_DWORD((in2 - low) / (high - low) * (_DWORD_TO_REAL(SHL(DWORD#2#1,_BYTE_TO_INT(bits))) - 1.0)   );
IF sx THEN Aout := SHL_DWORD(DWORD#2#1,_BYTE_TO_INT(sign)) OR Aout; END_IF;

(*
revision history

hm 18.1.2007		rev 1.1
	renamed Modul to aout.
	changed Output to 32 Bit max.
	corrected error with sign bit.

hm	13.9.2007		rev 1.2
	changed code to avoid warning under codesys 2.8.1

hm	2. dec 2007		rev 1.3
	changed code for better performance

hm	23. feb 2008	rev 1.4
	changed code for better performance
*)
(*@KEY@: END_WORKSHEET *)
END_FUNCTION

(* ---- AOUT1.ST ---- *)
(*@PROPERTIES_EX@
TYPE: POU
LOCALE: 0
IEC_LANGUAGE: ST
PLC_TYPE: independent
PROC_TYPE: independent
GROUP: ENGINEERING.SIGNAL_PROCESSING
*)
(*@KEY@:DESCRIPTION*)
version 1.0	23 feb 2008
programmer 	oscat
tested by	tobias

this module conditions an internal real value for a D/A converter.
(*@KEY@:END_DESCRIPTION*)
FUNCTION AOUT1:DWORD

(*Group:Default*)

VAR_INPUT
	IN :	REAL;
	BIT_0 :	INT;
	BIT_N :	INT;
	SIGN :	INT;
	LOW :	REAL;
	HIGH :	REAL;
END_VAR

VAR
	in2 :	REAL;
	sx :	BOOL;
END_VAR

(*@KEY@: WORKSHEET
NAME: AOUT1
IEC_LANGUAGE: ST
*)
(* if sign bit is defined *)

IF sign < 32 THEN
	sx := sign_R(in);
	in2 := ABS(in);
ELSE
    sx := FALSE;
	in2 := in;
END_IF;

(* begrenze in auf die zulässigen werte *)
in2 := LIMIT_REAL(low, in2, high);

(* Berechne den Ausgangswert *)
AOUT1 :=  SHL_DWORD(_REAL_TO_DWORD((in2 - low) / (high - low) * UDINT_TO_REAL(DWORD_TO_UDINT(SHL(DWORD#2#1,bit_n - Bit_0 + 1)) - UDINT#1)),Bit_0);

IF sx THEN AOUT1 := SHL(DWORD#2#1,sign) OR AOUT1; END_IF;

(* revision history
hm	23. feb 2008	rev 1.0
	original version

*)
(*@KEY@: END_WORKSHEET *)
END_FUNCTION

(* ---- CTRL_IN.ST ---- *)
(*@PROPERTIES_EX@
TYPE: POU
LOCALE: 0
IEC_LANGUAGE: ST
PLC_TYPE: independent
PROC_TYPE: independent
GROUP: ENGINEERING.CONTROL
*)
(*@KEY@:DESCRIPTION*)
version 1.0	2. jun 2008
programmer 	hugo
tested by	tobias
(*@KEY@:END_DESCRIPTION*)
FUNCTION CTRL_IN:REAL

(*Group:Default*)

VAR_INPUT
	SET_POINT :	REAL;
	ACTUAL :	REAL;
	NOISE :	REAL;
END_VAR

(*@KEY@: WORKSHEET
NAME: CTRL_IN
IEC_LANGUAGE: ST
*)
(* calculate the process error DIFF *)
CTRL_IN := DEAD_ZONE(SET_POINT - ACTUAL, NOISE);

(* revision history
hm 	2. jun. 2008 	rev 1.0
	original version

*)
(*@KEY@: END_WORKSHEET *)
END_FUNCTION

(* ---- DEC1.ST ---- *)
(*@PROPERTIES_EX@
TYPE: POU
LOCALE: 0
IEC_LANGUAGE: ST
PLC_TYPE: independent
PROC_TYPE: independent
GROUP: MATHEMATICAL.MATHE
*)
(*@KEY@:DESCRIPTION*)
version 1.1	27. oct. 2008
programmer 	hugo
tested by	oscat

This is a decrement function which decrements the variable X by 1 and if 0 is reached, it begins with M again.
_dec1(3,X) will generate 3,2,1,0,3,2,...
(*@KEY@:END_DESCRIPTION*)
FUNCTION DEC1:INT

(*Group:Default*)

VAR_INPUT
	X :	INT;
	N :	INT;
END_VAR

(*@KEY@: WORKSHEET
NAME: DEC1
IEC_LANGUAGE: ST
*)
IF X = 0 THEN
	DEC1 := N - 1;
ELSE
	DEC1 := X - 1;
END_IF;

(* this is a very elegant version but 50% slower
X := (X - 1 + N) MOD N;
*)

(* revision history
hm	13. oct. 2008	rev 1.0
	original version

hm	27. oct. 2008	rev 1.1
	added statement to return value for compatibility reasons
*)
(*@KEY@: END_WORKSHEET *)
END_FUNCTION

(* ---- FRMP_B.ST ---- *)
(*@PROPERTIES_EX@
TYPE: POU
LOCALE: 0
IEC_LANGUAGE: ST
PLC_TYPE: independent
PROC_TYPE: independent
GROUP: MATHEMATICAL.FUNCTIONS
*)
(*@KEY@:DESCRIPTION*)
version 1.0		17. feb. 2011
programmer 	    hugo
tested by		oscat

this function calculates a ramp and limits the output to 0 .. 255 without overflow problems

(*@KEY@:END_DESCRIPTION*)
FUNCTION FRMP_B:BYTE

(*Group:Default*)

VAR_INPUT
	START :	BYTE;
	DIR :	BOOL;
	TD :	TIME;
	TR :	TIME;
END_VAR

(*@KEY@: WORKSHEET
NAME: FRMP_B
IEC_LANGUAGE: ST
*)
IF TD < TR THEN
	FRMP_B := MIN(UDINT_TO_BYTE(DWORD_TO_UDINT(SHL(TIME_TO_DWORD(TD), 8)) / TIME_TO_UDINT(TR)), SEL(DIR, START, USINT_TO_BYTE(USINT#255 - BYTE_TO_USINT(START))));
	IF DIR THEN
		FRMP_B := USINT_TO_BYTE(BYTE_TO_USINT(START) + BYTE_TO_USINT(FRMP_B));
	ELSE
		FRMP_B := USINT_TO_BYTE(BYTE_TO_USINT(START) - BYTE_TO_USINT(FRMP_B));
	END_IF;
ELSE
	FRMP_B := SEL(DIR, BYTE#0, BYTE#255);
END_IF;

(* revision history

17. feb. 2011	rev 1.0
	new module

*)
(*@KEY@: END_WORKSHEET *)
END_FUNCTION

(* ---- INC.ST ---- *)
(*@PROPERTIES_EX@
TYPE: POU
LOCALE: 0
IEC_LANGUAGE: ST
PLC_TYPE: independent
PROC_TYPE: independent
GROUP: MATHEMATICAL.MATHE
*)
(*@KEY@:DESCRIPTION*)
version 1.1	15. jan 2008
programmer 	hugo
tested by	tobias

This is a increment function which increments the input X by the value D and compares the result with M.
if the output exceeds M it will continue to count from 0 again.
(*@KEY@:END_DESCRIPTION*)
FUNCTION INC:INT

(*Group:Default*)

VAR_INPUT
	X :	INT;
	D :	INT;
	M :	INT;
END_VAR

(*@KEY@: WORKSHEET
NAME: INC
IEC_LANGUAGE: ST
*)
inc := (X + D + M + 1) MOD (M + 1);

(* revision history
hm	7. feb 2007		REV 1.0
	original version

hm	15. jan 2008	rev 1.1
	allow for neagtive increment

*)
(*@KEY@: END_WORKSHEET *)
END_FUNCTION

(* ---- INC1.ST ---- *)
(*@PROPERTIES_EX@
TYPE: POU
LOCALE: 0
IEC_LANGUAGE: ST
PLC_TYPE: independent
PROC_TYPE: independent
GROUP: MATHEMATICAL.MATHE
*)
(*@KEY@:DESCRIPTION*)
version 1.2	23. feb. 2009
programmer 	hugo
tested by	oscat

This is a increment function which increments the variable X by 1 and if N is reached, it begins with 0 instead of N again.
inc1(X,3) will generate 0,1,2,0,1,.....
(*@KEY@:END_DESCRIPTION*)
FUNCTION INC1:INT

(*Group:Default*)

VAR_INPUT
	X :	INT;
	N :	INT;
END_VAR

(*@KEY@: WORKSHEET
NAME: INC1
IEC_LANGUAGE: ST
*)
IF X >= N - 1 THEN
	INC1 := 0;
ELSE
	INC1 := X + 1;
END_IF;

(* this elegant version is 50% slower
INC1 := X := (x + 1) MOD N;
*)

(* revision history
hm	13. oct. 2008	rev 1.0
	original version

hm	22. oct. 2008	rev 1.1
	added statement to return value for compatibility reasons

hm	23. feb. 2009	rev 1.2
 	when inc1 is called with X >= N inc will continue with 0
*)
(*@KEY@: END_WORKSHEET *)
END_FUNCTION

(* ---- INC2.ST ---- *)
(*@PROPERTIES_EX@
TYPE: POU
LOCALE: 0
IEC_LANGUAGE: ST
PLC_TYPE: independent
PROC_TYPE: independent
GROUP: MATHEMATICAL.MATHE
*)
(*@KEY@:DESCRIPTION*)
version 1.0	29. jun. 2008
programmer 	hugo
tested by	oscat

This function increments the input X by the value D and compares the result with U.
if the output exceeds U it will continue to count from L again.
(*@KEY@:END_DESCRIPTION*)
FUNCTION INC2:INT

(*Group:Default*)

VAR_INPUT
	X :	INT;
	D :	INT;
	L :	INT;
	U :	INT;
END_VAR

VAR
	tmp :	INT;
END_VAR

(*@KEY@: WORKSHEET
NAME: INC2
IEC_LANGUAGE: ST
*)
tmp := U - L + 1;
INC2 := (X + D - L + tmp) MOD tmp + L;

(* revision history
hm	29. jun. 2008		REV 1.0
	original version

*)
(*@KEY@: END_WORKSHEET *)
END_FUNCTION

(* ---- MANUAL.ST ---- *)
(*@PROPERTIES_EX@
TYPE: POU
LOCALE: 0
IEC_LANGUAGE: ST
PLC_TYPE: independent
PROC_TYPE: independent
GROUP: ENGINEERING.AUTOMATION
*)
(*@KEY@:DESCRIPTION*)
version 1.0	21. nov. 2008
programmer 	hugo
tested by	oscat

MANUAL is a manual override for digital signals.
when on and off = FALSE, the output follows IN.
ON = TRUE forces the output high, and OFF = TRUE forces the output low.
(*@KEY@:END_DESCRIPTION*)
FUNCTION MANUAL:BOOL

(*Group:Default*)

VAR_INPUT
	IN :	BOOL;
	ON :	BOOL;
	OFF :	BOOL;
END_VAR

(*@KEY@: WORKSHEET
NAME: MANUAL
IEC_LANGUAGE: ST
*)
MANUAL := NOT OFF AND (IN OR ON);

(* revision history
hm	21. nov 2008	rev 1.0
	original version

*)
(*@KEY@: END_WORKSHEET *)
END_FUNCTION

(* ---- SENSOR_INT.ST ---- *)
(*@PROPERTIES_EX@
TYPE: POU
LOCALE: 0
IEC_LANGUAGE: ST
PLC_TYPE: independent
PROC_TYPE: independent
GROUP: ENGINEERING.SENSOR
*)
(*@KEY@:DESCRIPTION*)
version 1.3	11. mar. 2009
programmer 	hugo
tested by	tobias

this function calculates the real resistance of a sensor RX given a parasitic resistor in parallel to the sensor and an additional serial resistor.
for example a parasitic parallel resistor for a PT100 can be ignored but a series resistor is the cable to the sensor.
for a humidity sensor, the parallel resistor is more dramatic and needs to be considered.
the function allows to consider a parallel and serial resistor at the same time.
with this function and known parasitic serial and parallel resistors the true resistance of the sensor can be calculated.

(*@KEY@:END_DESCRIPTION*)
FUNCTION SENSOR_INT:REAL

(*Group:Default*)

VAR_INPUT
	VOLTAGE :	REAL;
	CURRENT :	REAL;
	RP :	REAL;
	RS :	REAL;
END_VAR

VAR
	RG :	REAL;
END_VAR

(*@KEY@: WORKSHEET
NAME: SENSOR_INT
IEC_LANGUAGE: ST
*)
IF current <> 0.0 THEN
	RG := voltage / current;
	SENSOR_INT := RP * ( RG - RS) / ( RP + RS - RG);
END_IF;

(* revisaion history

hm 20.1.2007		rev 1.1
	deleted input R0 which was not needed.

hm	2. dec 2007	rev 1.2
	corrected an error in formula and improoved speed

hm	11. mar. 2009	rev 1.3
	changed real constants to use dot syntax

*)
(*@KEY@: END_WORKSHEET *)
END_FUNCTION

(* ---- STAIR.ST ---- *)
(*@PROPERTIES_EX@
TYPE: POU
LOCALE: 0
IEC_LANGUAGE: ST
PLC_TYPE: independent
PROC_TYPE: independent
GROUP: ENGINEERING.SIGNAL_PROCESSING
*)
(*@KEY@:DESCRIPTION*)
version 1.4	10. mar. 2009
programmer 	oscat
tested by	tobias

the function stair converts an anlog input signal to a staircase like output.
D is the step width for the output signal.
if D = 0 then the output follows the input without a chage.
(*@KEY@:END_DESCRIPTION*)
FUNCTION STAIR:REAL

(*Group:Default*)

VAR_INPUT
	X :	REAL;
	D :	REAL;
END_VAR

(*@KEY@: WORKSHEET
NAME: STAIR
IEC_LANGUAGE: ST
*)
IF D > 0.0 THEN
	STAIR := DINT_TO_REAL(_REAL_TO_DINT(X / D)) * D;
ELSE
	STAIR := X;
END_IF;

(* revision history
hm	28 jan 2007		rev 1.0
	original version

hm	27 dec 2007		rev 1.1
	changed code for better performance

hm	6. jan 2008		rev 1.2
	further performance improvement

hm	26. oct. 2008		rev 1.3
	optimized code

hm	10. mar. 2009	rev 1.4
	real constants updated to new systax using dot

*)
(*@KEY@: END_WORKSHEET *)
END_FUNCTION

(* ---- TIMECHECK.ST ---- *)
(*@PROPERTIES_EX@
TYPE: POU
LOCALE: 0
IEC_LANGUAGE: ST
PLC_TYPE: independent
PROC_TYPE: independent
GROUP: TIME_DATE
*)
(*@KEY@:DESCRIPTION*)
version 1.0	19. jul. 2009
programmer 	oscat
tested by	oscat

this function retruns true if the daytime TD is between start and stop and returns true if so.
if you want to generate an event to span over midnight, start timemust be later than the stop time.

(*@KEY@:END_DESCRIPTION*)
FUNCTION TIMECHECK:BOOL

(*Group:Default*)

VAR_INPUT
	TD :	UDINT;
	START :	UDINT;
	STOP :	UDINT;
END_VAR

(*@KEY@: WORKSHEET
NAME: TIMECHECK
IEC_LANGUAGE: ST
*)
IF stop < start THEN
	TIMECHECK := start <= TD OR  TD < stop;
ELSE
	TIMECHECK := start <= TD AND TD < stop;
END_IF;

(* revision history
hm 19. jul. 2009	rev 1.0
	original release

*)
(*@KEY@: END_WORKSHEET *)
END_FUNCTION
